RoboDK station: Conveyor_Station.rdk

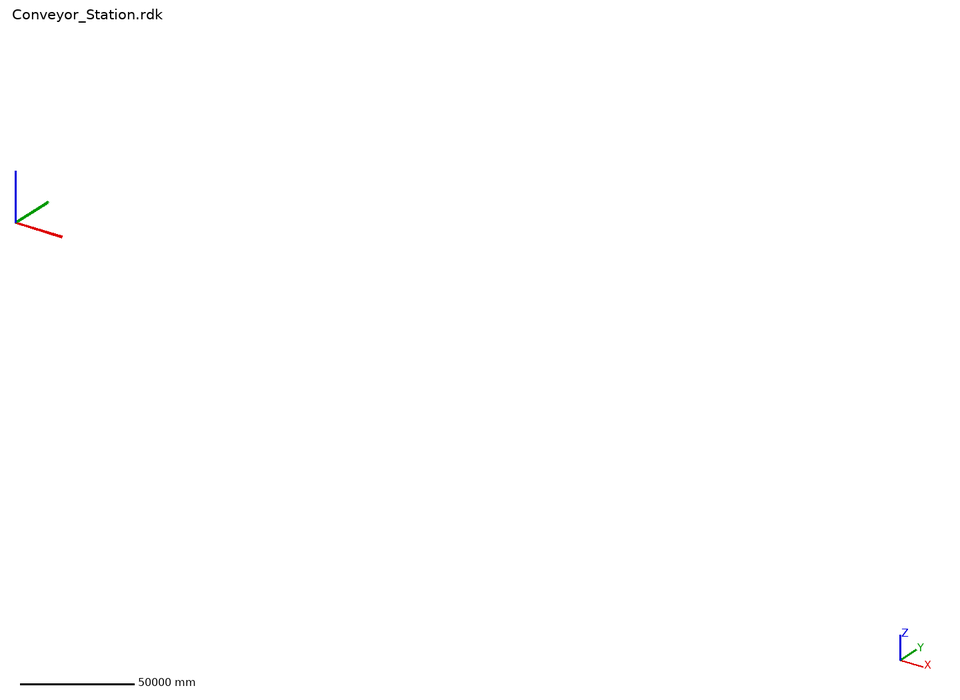
[picture v0: the station drawn from its stored meshes, robots at their saved joint values, targets as dots, program paths as lines]
Station Conveyor_Station (saved by RoboDK 6.0.1). Poses are relative to the parent item; angles as X-Y-Z fixed-axis rotations.
  - frame Conveyor Belt Wide (2m) Base at (0, 0, 0) mm
    - robot Conveyor Belt Wide (2m): 1 axes
        modified DH rows (alpha deg, a mm, theta deg, d mm): 0, 0, 0, 0 linear
        base shift (0, 0, 0) mm, rotated rx 0 ry 90 rz 0 deg
        joint limits [-900000] to [900000]; home [0]; saved at [-400005]
      - frame Conveyor Frame at (0, 0, 0) mm
        - object Box at (896234, 103.35, 13.17) mm, rotated rx -0.5 ry 0.31 rz 13.64 deg, size 10 x 20 x 5 mm, geometry from box.sld
        - object Box at (895766, 103.35, 13.17) mm, rotated rx -0.51 ry 0.3 rz 12.18 deg, size 10 x 20 x 5 mm, geometry from box.sld
        - object Box at (895300, 103.35, 13.17) mm, rotated rx -0.59 ry -0.09 rz -27.08 deg, size 10 x 20 x 5 mm, geometry from box.sld
        - object Box at (894830, 103.35, 13.17) mm, rotated rx -0.59 ry 0.03 rz -14.87 deg, size 10 x 20 x 5 mm, geometry from box.sld
        - object Box at (894363, 103.35, 13.17) mm, rotated rx -0.59 ry 0.08 rz -10.87 deg, size 10 x 20 x 5 mm, geometry from box.sld
        - object Box at (893893, 103.35, 13.17) mm, rotated rx -0.54 ry -0.25 rz -42.71 deg, size 10 x 20 x 5 mm, geometry from box.sld
        - object Box at (893423, 103.35, 13.17) mm, rotated rx -0.58 ry -0.12 rz -29.69 deg, size 10 x 20 x 5 mm, geometry from box.sld
        - object Box at (892951, 103.35, 13.17) mm, rotated rx -0.54 ry -0.25 rz -42.74 deg, size 10 x 20 x 5 mm, geometry from box.sld
        - object Box at (892481, 103.35, 13.17) mm, rotated rx -0.56 ry -0.19 rz -36.39 deg, size 10 x 20 x 5 mm, geometry from box.sld
        - object Box at (892010, 103.35, 13.17) mm, rotated rx -0.38 ry 0.45 rz 31.55 deg, size 10 x 20 x 5 mm, geometry from box.sld
        - object Box at (891537, 103.35, 13.17) mm, rotated rx -0.58 ry -0.14 rz -31.84 deg, size 10 x 20 x 5 mm, geometry from box.sld
        - object Box at (891061, 103.35, 13.17) mm, rotated rx -0.45 ry 0.39 rz 23.02 deg, size 10 x 20 x 5 mm, geometry from box.sld
        - object Box at (889213, 103.35, 13.17) mm, rotated rx -0.58 ry 0.14 rz -4.6 deg, size 10 x 20 x 5 mm, geometry from box.sld
        - object Box at (887815, 103.35, 13.17) mm, rotated rx -0.5 ry 0.33 rz 15.16 deg, size 10 x 20 x 5 mm, geometry from box.sld
        - object Box at (884546, 103.35, 13.17) mm, rotated rx -0.51 ry 0.31 rz 13.23 deg, size 10 x 20 x 5 mm, geometry from box.sld
        - object Box at (884069, 103.35, 13.17) mm, rotated rx -0.53 ry -0.27 rz -44.95 deg, size 10 x 20 x 5 mm, geometry from box.sld
        - object Box at (883940, 103.35, 13.17) mm, rotated rx -0.42 ry 0.42 rz 26.41 deg, size 10 x 20 x 5 mm, geometry from box.sld
        - object Box at (883628, 103.35, 13.17) mm, rotated rx -0.43 ry 0.41 rz 25.46 deg, size 10 x 20 x 5 mm, geometry from box.sld
        - object Box at (881822, 103.35, 13.17) mm, rotated rx -0.29 ry 0.52 rz 42.29 deg, size 10 x 20 x 5 mm, geometry from box.sld
        - object Box at (881392, 103.35, 13.17) mm, rotated rx -0.58 ry 0.12 rz -6.43 deg, size 10 x 20 x 5 mm, geometry from box.sld
        - object Box at (880938, 103.35, 13.17) mm, rotated rx -0.33 ry 0.5 rz 38.54 deg, size 10 x 20 x 5 mm, geometry from box.sld
        - object Box at (880498, 103.35, 13.17) mm, rotated rx -0.44 ry 0.4 rz 23.86 deg, size 10 x 20 x 5 mm, geometry from box.sld
        - object Box at (880042, 103.35, 13.17) mm, rotated rx -0.58 ry 0.13 rz -5.68 deg, size 10 x 20 x 5 mm, geometry from box.sld
        - object Box at (879599, 103.35, 13.17) mm, rotated rx -0.55 ry 0.22 rz 3.99 deg, size 10 x 20 x 5 mm, geometry from box.sld
        - object Box at (879164, 103.35, 13.17) mm, rotated rx -0.59 ry -0.01 rz -18.88 deg, size 10 x 20 x 5 mm, geometry from box.sld
        - object Box at (878722, 103.35, 13.17) mm, rotated rx -0.54 ry -0.24 rz -41.68 deg, size 10 x 20 x 5 mm, geometry from box.sld
        - object Box at (878276, 103.35, 13.17) mm, rotated rx -0.43 ry 0.41 rz 25.6 deg, size 10 x 20 x 5 mm, geometry from box.sld
        - object Box at (877829, 103.35, 13.17) mm, rotated rx -0.55 ry 0.23 rz 4.27 deg, size 10 x 20 x 5 mm, geometry from box.sld
        - object Box at (877389, 103.35, 13.17) mm, rotated rx -0.49 ry 0.33 rz 16.13 deg, size 10 x 20 x 5 mm, geometry from box.sld
        - object Box at (876944, 103.35, 13.17) mm, rotated rx -0.5 ry 0.33 rz 15.3 deg, size 10 x 20 x 5 mm, geometry from box.sld
        - object Box at (876499, 103.35, 13.17) mm, rotated rx -0.33 ry 0.5 rz 38.6 deg, size 10 x 20 x 5 mm, geometry from box.sld
        - object Box at (876043, 103.35, 13.17) mm, rotated rx -0.41 ry 0.43 rz 28.42 deg, size 10 x 20 x 5 mm, geometry from box.sld
        - object Box at (875592, 103.35, 13.17) mm, rotated rx -0.59 ry 0.03 rz -15.71 deg, size 10 x 20 x 5 mm, geometry from box.sld
        - object Box at (867999, 103.35, 13.17) mm, rotated rx -0.55 ry -0.22 rz -39.96 deg, size 10 x 20 x 5 mm, geometry from box.sld
        - object Box at (867540, 103.35, 13.17) mm, rotated rx -0.43 ry 0.41 rz 25.54 deg, size 10 x 20 x 5 mm, geometry from box.sld
        - object Box at (867083, 103.35, 13.17) mm, rotated rx -0.55 ry 0.23 rz 5.04 deg, size 10 x 20 x 5 mm, geometry from box.sld
        - object Box at (866626, 103.35, 13.17) mm, rotated rx -0.53 ry 0.26 rz 7.77 deg, size 10 x 20 x 5 mm, geometry from box.sld
        - object Box at (866172, 103.35, 13.17) mm, rotated rx -0.59 ry 0.09 rz -9.75 deg, size 10 x 20 x 5 mm, geometry from box.sld
        - object Box at (865727, 103.35, 13.17) mm, rotated rx -0.51 ry 0.31 rz 13.25 deg, size 10 x 20 x 5 mm, geometry from box.sld
        - object Box at (865279, 103.35, 13.17) mm, rotated rx -0.54 ry 0.24 rz 5.36 deg, size 10 x 20 x 5 mm, geometry from box.sld
        - object Box at (864826, 103.35, 13.17) mm, rotated rx -0.55 ry 0.23 rz 4.39 deg, size 10 x 20 x 5 mm, geometry from box.sld
        - object Box at (864371, 103.35, 13.17) mm, rotated rx -0.4 ry 0.44 rz 29 deg, size 10 x 20 x 5 mm, geometry from box.sld
        - object Box at (863914, 103.35, 13.17) mm, rotated rx -0.59 ry 0.09 rz -9.63 deg, size 10 x 20 x 5 mm, geometry from box.sld
        - object Box at (863455, 103.35, 13.17) mm, rotated rx -0.55 ry -0.22 rz -39.93 deg, size 10 x 20 x 5 mm, geometry from box.sld
        - object Box at (862988, 103.35, 13.17) mm, rotated rx -0.37 ry 0.46 rz 33.18 deg, size 10 x 20 x 5 mm, geometry from box.sld
        - object Box at (862512, 103.35, 13.17) mm, rotated rx -0.42 ry 0.42 rz 26.7 deg, size 10 x 20 x 5 mm, geometry from box.sld
        - object Box at (862049, 103.35, 13.17) mm, rotated rx -0.59 ry -0.07 rz -25.35 deg, size 10 x 20 x 5 mm, geometry from box.sld
        - object Box at (861585, 103.35, 13.17) mm, rotated rx -0.58 ry -0.13 rz -30.37 deg, size 10 x 20 x 5 mm, geometry from box.sld
        - object Box at (861121, 103.35, 13.17) mm, rotated rx -0.48 ry 0.35 rz 17.4 deg, size 10 x 20 x 5 mm, geometry from box.sld
        - object Box at (860654, 103.35, 13.17) mm, rotated rx -0.3 ry 0.51 rz 41.14 deg, size 10 x 20 x 5 mm, geometry from box.sld
        - object Box at (860190, 103.35, 13.17) mm, rotated rx -0.56 ry 0.2 rz 1.9 deg, size 10 x 20 x 5 mm, geometry from box.sld
        - object Box at (859725, 103.35, 13.17) mm, rotated rx -0.56 ry -0.21 rz -38.78 deg, size 10 x 20 x 5 mm, geometry from box.sld
        - object Box at (859255, 103.35, 13.17) mm, rotated rx -0.54 ry -0.25 rz -42.79 deg, size 10 x 20 x 5 mm, geometry from box.sld
        - object Box at (858791, 103.35, 13.17) mm, rotated rx -0.45 ry 0.38 rz 21.87 deg, size 10 x 20 x 5 mm, geometry from box.sld
        - object Box at (858319, 103.35, 13.17) mm, rotated rx -0.56 ry -0.21 rz -38.56 deg, size 10 x 20 x 5 mm, geometry from box.sld
        - object Box at (857850, 103.35, 13.17) mm, rotated rx -0.59 ry 0.09 rz -9.73 deg, size 10 x 20 x 5 mm, geometry from box.sld
        - object Box at (857380, 103.35, 13.17) mm, rotated rx -0.51 ry 0.31 rz 13.08 deg, size 10 x 20 x 5 mm, geometry from box.sld
        - object Box at (856914, 103.35, 13.17) mm, rotated rx -0.57 ry 0.16 rz -2.36 deg, size 10 x 20 x 5 mm, geometry from box.sld
        - object Box at (856441, 103.35, 13.17) mm, rotated rx -0.55 ry 0.23 rz 4.5 deg, size 10 x 20 x 5 mm, geometry from box.sld
        - object Box at (855972, 103.35, 13.17) mm, rotated rx -0.58 ry 0.13 rz -5.45 deg, size 10 x 20 x 5 mm, geometry from box.sld
        - object Box at (855499, 103.35, 13.17) mm, rotated rx -0.28 ry 0.52 rz 43.43 deg, size 10 x 20 x 5 mm, geometry from box.sld
        - object Box at (855027, 103.35, 13.17) mm, rotated rx -0.54 ry -0.24 rz -42.08 deg, size 10 x 20 x 5 mm, geometry from box.sld
        - object Box at (854558, 103.35, 13.17) mm, rotated rx -0.58 ry -0.12 rz -30.27 deg, size 10 x 20 x 5 mm, geometry from box.sld
        - object Box at (854093, 103.35, 13.17) mm, rotated rx -0.46 ry 0.37 rz 20.93 deg, size 10 x 20 x 5 mm, geometry from box.sld
        - object Box at (853622, 103.35, 13.17) mm, rotated rx -0.55 ry 0.23 rz 4.81 deg, size 10 x 20 x 5 mm, geometry from box.sld
        - object Box at (853148, 103.35, 13.17) mm, rotated rx -0.4 ry 0.44 rz 29.12 deg, size 10 x 20 x 5 mm, geometry from box.sld
        - object Box at (852676, 103.35, 13.17) mm, rotated rx -0.58 ry 0.14 rz -4.4 deg, size 10 x 20 x 5 mm, geometry from box.sld
        - object Box at (852209, 103.35, 13.17) mm, rotated rx -0.55 ry -0.22 rz -39.44 deg, size 10 x 20 x 5 mm, geometry from box.sld
        - object Box at (851737, 103.35, 13.17) mm, rotated rx -0.48 ry 0.35 rz 18.04 deg, size 10 x 20 x 5 mm, geometry from box.sld
        - object Box at (851258, 103.35, 13.17) mm, rotated rx -0.56 ry 0.2 rz 1.49 deg, size 10 x 20 x 5 mm, geometry from box.sld
        - object Box at (850779, 103.35, 13.17) mm, rotated rx -0.59 ry -0.05 rz -22.99 deg, size 10 x 20 x 5 mm, geometry from box.sld
        - object Box at (850302, 103.35, 13.17) mm, rotated rx -0.58 ry -0.14 rz -32.02 deg, size 10 x 20 x 5 mm, geometry from box.sld
        - object Box at (849825, 103.35, 13.17) mm, rotated rx -0.53 ry 0.27 rz 9.09 deg, size 10 x 20 x 5 mm, geometry from box.sld
        - object Box at (849347, 103.35, 13.17) mm, rotated rx -0.58 ry 0.1 rz -8 deg, size 10 x 20 x 5 mm, geometry from box.sld
        - object Box at (848871, 103.35, 13.17) mm, rotated rx -0.29 ry 0.52 rz 42.76 deg, size 10 x 20 x 5 mm, geometry from box.sld
        - object Box at (848385, 103.35, 13.17) mm, rotated rx -0.32 ry 0.5 rz 39.44 deg, size 10 x 20 x 5 mm, geometry from box.sld
        - object Box at (847911, 103.35, 13.17) mm, rotated rx -0.54 ry 0.24 rz 6.18 deg, size 10 x 20 x 5 mm, geometry from box.sld
        - object Box at (847434, 103.35, 13.17) mm, rotated rx -0.53 ry 0.27 rz 8.37 deg, size 10 x 20 x 5 mm, geometry from box.sld
        - object Box at (846952, 103.35, 13.17) mm, rotated rx -0.55 ry 0.21 rz 2.67 deg, size 10 x 20 x 5 mm, geometry from box.sld
        - object Box at (846476, 103.35, 13.17) mm, rotated rx -0.47 ry 0.36 rz 19.66 deg, size 10 x 20 x 5 mm, geometry from box.sld
        - object Box at (845998, 103.35, 13.17) mm, rotated rx -0.32 ry 0.5 rz 39.15 deg, size 10 x 20 x 5 mm, geometry from box.sld
        - object Box at (845516, 103.35, 13.17) mm, rotated rx -0.57 ry 0.18 rz -0.46 deg, size 10 x 20 x 5 mm, geometry from box.sld
        - object Box at (845034, 103.35, 13.17) mm, rotated rx -0.59 ry -0.04 rz -21.91 deg, size 10 x 20 x 5 mm, geometry from box.sld
        - object Box at (844553, 103.35, 13.17) mm, rotated rx -0.59 ry -0.09 rz -26.83 deg, size 10 x 20 x 5 mm, geometry from box.sld
        - object Box at (844070, 103.35, 13.17) mm, rotated rx -0.59 ry -0.01 rz -19.02 deg, size 10 x 20 x 5 mm, geometry from box.sld
        - object Box at (843586, 103.35, 13.17) mm, rotated rx -0.59 ry -0.08 rz -25.81 deg, size 10 x 20 x 5 mm, geometry from box.sld
        - object Box at (843104, 103.35, 13.17) mm, rotated rx -0.59 ry -0.01 rz -19.6 deg, size 10 x 20 x 5 mm, geometry from box.sld
        - object Box at (842621, 103.35, 13.17) mm, rotated rx -0.38 ry 0.45 rz 31.78 deg, size 10 x 20 x 5 mm, geometry from box.sld
        - object Box at (842135, 103.35, 13.17) mm, rotated rx -0.55 ry -0.23 rz -40.91 deg, size 10 x 20 x 5 mm, geometry from box.sld
        - object Box at (841652, 103.35, 13.17) mm, rotated rx -0.59 ry -0.05 rz -22.69 deg, size 10 x 20 x 5 mm, geometry from box.sld
        - object Box at (841168, 103.35, 13.17) mm, rotated rx -0.54 ry -0.26 rz -43.77 deg, size 10 x 20 x 5 mm, geometry from box.sld
        - object Box at (840683, 103.35, 13.17) mm, rotated rx -0.39 ry 0.45 rz 30.57 deg, size 10 x 20 x 5 mm, geometry from box.sld
        - object Box at (840198, 103.35, 13.17) mm, rotated rx -0.57 ry -0.16 rz -33.5 deg, size 10 x 20 x 5 mm, geometry from box.sld
        - object Box at (839715, 103.35, 13.17) mm, rotated rx -0.58 ry -0.12 rz -30.28 deg, size 10 x 20 x 5 mm, geometry from box.sld
        - object Box at (839227, 103.35, 13.17) mm, rotated rx -0.35 ry 0.48 rz 35.52 deg, size 10 x 20 x 5 mm, geometry from box.sld
        - object Box at (838741, 103.35, 13.17) mm, rotated rx -0.58 ry 0.1 rz -8.02 deg, size 10 x 20 x 5 mm, geometry from box.sld
        - object Box at (838251, 103.35, 13.17) mm, rotated rx -0.57 ry -0.15 rz -33.01 deg, size 10 x 20 x 5 mm, geometry from box.sld
        - object Box at (837766, 103.35, 13.17) mm, rotated rx -0.47 ry 0.36 rz 19.31 deg, size 10 x 20 x 5 mm, geometry from box.sld
        - object Box at (837279, 103.35, 13.17) mm, rotated rx -0.57 ry 0.15 rz -3.62 deg, size 10 x 20 x 5 mm, geometry from box.sld
        - object Box at (836786, 103.35, 13.17) mm, rotated rx -0.3 ry 0.51 rz 41.2 deg, size 10 x 20 x 5 mm, geometry from box.sld
        - object Box at (836295, 103.35, 13.17) mm, rotated rx -0.35 ry 0.48 rz 35.79 deg, size 10 x 20 x 5 mm, geometry from box.sld
        - object Box at (835805, 103.35, 13.17) mm, rotated rx -0.58 ry 0.11 rz -7.26 deg, size 10 x 20 x 5 mm, geometry from box.sld
        - object Box at (835317, 103.35, 13.17) mm, rotated rx -0.58 ry 0.14 rz -4.75 deg, size 10 x 20 x 5 mm, geometry from box.sld
        - object Box at (834829, 103.35, 13.17) mm, rotated rx -0.48 ry 0.35 rz 18.31 deg, size 10 x 20 x 5 mm, geometry from box.sld
        - object Box at (834338, 103.35, 13.17) mm, rotated rx -0.44 ry 0.4 rz 24.11 deg, size 10 x 20 x 5 mm, geometry from box.sld
        - object Box at (833842, 103.35, 13.17) mm, rotated rx -0.55 ry -0.22 rz -39.64 deg, size 10 x 20 x 5 mm, geometry from box.sld
        - object Box at (833349, 103.35, 13.17) mm, rotated rx -0.46 ry 0.37 rz 20.57 deg, size 10 x 20 x 5 mm, geometry from box.sld
        - object Box at (832860, 103.35, 13.17) mm, rotated rx -0.55 ry -0.23 rz -40.82 deg, size 10 x 20 x 5 mm, geometry from box.sld
        - object Box at (832363, 103.35, 13.17) mm, rotated rx -0.58 ry 0.1 rz -8.13 deg, size 10 x 20 x 5 mm, geometry from box.sld
        - object Box at (831873, 103.35, 13.17) mm, rotated rx -0.59 ry -0.08 rz -26.3 deg, size 10 x 20 x 5 mm, geometry from box.sld
        - object Box at (831377, 103.35, 13.17) mm, rotated rx -0.52 ry 0.28 rz 10.12 deg, size 10 x 20 x 5 mm, geometry from box.sld
        - object Box at (830887, 103.35, 13.17) mm, rotated rx -0.59 ry 0.02 rz -16.15 deg, size 10 x 20 x 5 mm, geometry from box.sld
        - object Box at (830394, 103.35, 13.17) mm, rotated rx -0.59 ry -0.03 rz -21.06 deg, size 10 x 20 x 5 mm, geometry from box.sld
        - object Box at (829901, 103.35, 13.17) mm, rotated rx -0.59 ry -0.02 rz -20.25 deg, size 10 x 20 x 5 mm, geometry from box.sld
        - object Box at (829404, 103.35, 13.17) mm, rotated rx -0.49 ry 0.34 rz 17.03 deg, size 10 x 20 x 5 mm, geometry from box.sld
        - object Box at (828911, 103.35, 13.17) mm, rotated rx -0.56 ry 0.19 rz 0.53 deg, size 10 x 20 x 5 mm, geometry from box.sld
        - object Box at (828417, 103.35, 13.17) mm, rotated rx -0.32 ry 0.5 rz 38.99 deg, size 10 x 20 x 5 mm, geometry from box.sld
        - object Box at (827919, 103.35, 13.17) mm, rotated rx -0.58 ry -0.14 rz -31.79 deg, size 10 x 20 x 5 mm, geometry from box.sld
        - object Box at (827419, 103.35, 13.17) mm, rotated rx -0.47 ry 0.36 rz 19.71 deg, size 10 x 20 x 5 mm, geometry from box.sld
        - object Box at (826919, 103.35, 13.17) mm, rotated rx -0.28 ry 0.52 rz 43.35 deg, size 10 x 20 x 5 mm, geometry from box.sld
        - object Box at (826422, 103.35, 13.17) mm, rotated rx -0.47 ry 0.37 rz 20.05 deg, size 10 x 20 x 5 mm, geometry from box.sld
        - object Box at (825923, 103.35, 13.17) mm, rotated rx -0.59 ry -0.09 rz -27.23 deg, size 10 x 20 x 5 mm, geometry from box.sld
        - object Box at (825422, 103.35, 13.17) mm, rotated rx -0.59 ry -0.02 rz -20.55 deg, size 10 x 20 x 5 mm, geometry from box.sld
        - object Box at (824929, 103.35, 13.17) mm, rotated rx -0.54 ry 0.25 rz 6.23 deg, size 10 x 20 x 5 mm, geometry from box.sld
        - object Box at (824425, 103.35, 13.17) mm, rotated rx -0.59 ry 0 rz -17.98 deg, size 10 x 20 x 5 mm, geometry from box.sld
        - object Box at (823928, 103.35, 13.17) mm, rotated rx -0.31 ry 0.5 rz 39.89 deg, size 10 x 20 x 5 mm, geometry from box.sld
        - object Box at (823424, 103.35, 13.17) mm, rotated rx -0.55 ry 0.23 rz 4.6 deg, size 10 x 20 x 5 mm, geometry from box.sld
        - object Box at (822920, 103.35, 13.17) mm, rotated rx -0.4 ry 0.44 rz 29.82 deg, size 10 x 20 x 5 mm, geometry from box.sld
        - object Box at (822418, 103.35, 13.17) mm, rotated rx -0.34 ry 0.49 rz 36.72 deg, size 10 x 20 x 5 mm, geometry from box.sld
        - object Box at (821917, 103.35, 13.17) mm, rotated rx -0.58 ry -0.12 rz -30.21 deg, size 10 x 20 x 5 mm, geometry from box.sld
        - object Box at (821420, 103.35, 13.17) mm, rotated rx -0.59 ry 0.04 rz -14.15 deg, size 10 x 20 x 5 mm, geometry from box.sld
        - object Box at (820919, 103.35, 13.17) mm, rotated rx -0.59 ry -0.08 rz -25.75 deg, size 10 x 20 x 5 mm, geometry from box.sld
        - object Box at (820410, 103.35, 13.17) mm, rotated rx -0.5 ry 0.33 rz 15.32 deg, size 10 x 20 x 5 mm, geometry from box.sld
        - object Box at (819909, 103.35, 13.17) mm, rotated rx -0.53 ry 0.26 rz 7.55 deg, size 10 x 20 x 5 mm, geometry from box.sld
        - object Box at (819403, 103.35, 13.17) mm, rotated rx -0.28 ry 0.52 rz 43.76 deg, size 10 x 20 x 5 mm, geometry from box.sld
        - object Box at (818898, 103.35, 13.17) mm, rotated rx -0.55 ry 0.21 rz 2.65 deg, size 10 x 20 x 5 mm, geometry from box.sld
        - object Box at (818392, 103.35, 13.17) mm, rotated rx -0.32 ry 0.5 rz 39.41 deg, size 10 x 20 x 5 mm, geometry from box.sld
        - object Box at (817887, 103.35, 13.17) mm, rotated rx -0.33 ry 0.49 rz 38.25 deg, size 10 x 20 x 5 mm, geometry from box.sld
        - object Box at (817383, 103.35, 13.17) mm, rotated rx -0.58 ry -0.11 rz -28.6 deg, size 10 x 20 x 5 mm, geometry from box.sld
        - object Box at (816879, 103.35, 13.17) mm, rotated rx -0.38 ry 0.46 rz 31.95 deg, size 10 x 20 x 5 mm, geometry from box.sld
        - object Box at (816374, 103.35, 13.17) mm, rotated rx -0.3 ry 0.51 rz 41.87 deg, size 10 x 20 x 5 mm, geometry from box.sld
        - object Box at (815868, 103.35, 13.17) mm, rotated rx -0.28 ry 0.52 rz 44.01 deg, size 10 x 20 x 5 mm, geometry from box.sld
        - object Box at (815360, 103.35, 13.17) mm, rotated rx -0.37 ry 0.46 rz 32.8 deg, size 10 x 20 x 5 mm, geometry from box.sld
        - object Box at (814853, 103.35, 13.17) mm, rotated rx -0.59 ry 0.07 rz -11.65 deg, size 10 x 20 x 5 mm, geometry from box.sld
        - object Box at (814348, 103.35, 13.17) mm, rotated rx -0.59 ry 0 rz -18.55 deg, size 10 x 20 x 5 mm, geometry from box.sld
        - object Box at (813832, 103.35, 13.17) mm, rotated rx -0.44 ry 0.4 rz 24.43 deg, size 10 x 20 x 5 mm, geometry from box.sld
        - object Box at (813321, 103.35, 13.17) mm, rotated rx -0.51 ry 0.31 rz 13.24 deg, size 10 x 20 x 5 mm, geometry from box.sld
        - object Box at (812812, 103.35, 13.17) mm, rotated rx -0.41 ry 0.43 rz 28.3 deg, size 10 x 20 x 5 mm, geometry from box.sld
        - object Box at (812298, 103.35, 13.17) mm, rotated rx -0.27 ry 0.53 rz 44.37 deg, size 10 x 20 x 5 mm, geometry from box.sld
        - object Box at (811784, 103.35, 13.17) mm, rotated rx -0.5 ry 0.32 rz 13.91 deg, size 10 x 20 x 5 mm, geometry from box.sld
        - object Box at (811274, 103.35, 13.17) mm, rotated rx -0.59 ry -0.02 rz -20.03 deg, size 10 x 20 x 5 mm, geometry from box.sld
        - object Box at (810763, 103.35, 13.17) mm, rotated rx -0.59 ry -0.02 rz -19.79 deg, size 10 x 20 x 5 mm, geometry from box.sld
        - object Box at (810254, 103.35, 13.17) mm, rotated rx -0.35 ry 0.48 rz 35.74 deg, size 10 x 20 x 5 mm, geometry from box.sld
        - object Box at (809736, 103.35, 13.17) mm, rotated rx -0.59 ry 0.09 rz -9.12 deg, size 10 x 20 x 5 mm, geometry from box.sld
        - object Box at (809227, 103.35, 13.17) mm, rotated rx -0.56 ry 0.19 rz 0.29 deg, size 10 x 20 x 5 mm, geometry from box.sld
        - object Box at (808709, 103.35, 13.17) mm, rotated rx -0.38 ry 0.45 rz 31.82 deg, size 10 x 20 x 5 mm, geometry from box.sld
        - object Box at (808195, 103.35, 13.17) mm, rotated rx -0.4 ry 0.44 rz 29.46 deg, size 10 x 20 x 5 mm, geometry from box.sld
        - object Box at (807680, 103.35, 13.17) mm, rotated rx -0.53 ry 0.26 rz 7.88 deg, size 10 x 20 x 5 mm, geometry from box.sld
        - object Box at (807162, 103.35, 13.17) mm, rotated rx -0.51 ry 0.3 rz 12.3 deg, size 10 x 20 x 5 mm, geometry from box.sld
        - object Box at (806641, 103.35, 13.17) mm, rotated rx -0.3 ry 0.51 rz 41.63 deg, size 10 x 20 x 5 mm, geometry from box.sld
        - object Box at (806130, 103.35, 13.17) mm, rotated rx -0.56 ry 0.19 rz 0.61 deg, size 10 x 20 x 5 mm, geometry from box.sld
        - object Box at (805613, 103.35, 13.17) mm, rotated rx -0.45 ry 0.39 rz 22.73 deg, size 10 x 20 x 5 mm, geometry from box.sld
        - object Box at (805094, 103.35, 13.17) mm, rotated rx -0.59 ry -0.03 rz -20.82 deg, size 10 x 20 x 5 mm, geometry from box.sld
        - object Box at (804579, 103.35, 13.17) mm, rotated rx -0.55 ry -0.22 rz -40.13 deg, size 10 x 20 x 5 mm, geometry from box.sld
        - object Box at (804064, 103.35, 13.17) mm, rotated rx -0.58 ry 0.13 rz -5.18 deg, size 10 x 20 x 5 mm, geometry from box.sld
        - object Box at (803548, 103.35, 13.17) mm, rotated rx -0.55 ry 0.21 rz 2.72 deg, size 10 x 20 x 5 mm, geometry from box.sld
        - object Box at (803030, 103.35, 13.17) mm, rotated rx -0.36 ry 0.47 rz 34.01 deg, size 10 x 20 x 5 mm, geometry from box.sld
        - object Box at (802512, 103.35, 13.17) mm, rotated rx -0.51 ry 0.3 rz 11.68 deg, size 10 x 20 x 5 mm, geometry from box.sld
        - object Box at (801994, 103.35, 13.17) mm, rotated rx -0.57 ry -0.17 rz -34.33 deg, size 10 x 20 x 5 mm, geometry from box.sld
        - object Box at (801472, 103.35, 13.17) mm, rotated rx -0.5 ry 0.32 rz 14.1 deg, size 10 x 20 x 5 mm, geometry from box.sld
        - object Box at (800951, 103.35, 13.17) mm, rotated rx -0.51 ry 0.31 rz 13.06 deg, size 10 x 20 x 5 mm, geometry from box.sld
        - object Box at (800432, 103.35, 13.17) mm, rotated rx -0.59 ry -0.02 rz -20.34 deg, size 10 x 20 x 5 mm, geometry from box.sld
        - object Box at (800001, 103.35, 13.17) mm, rotated rx -0.59 ry 0.03 rz -15.33 deg, size 10 x 20 x 5 mm, geometry from box.sld
        - object Box at (799501, 103.35, 13.17) mm, rotated rx -0.54 ry -0.25 rz -43.39 deg, size 10 x 20 x 5 mm, geometry from box.sld
        - object Box at (798979, 103.35, 13.17) mm, rotated rx -0.4 ry 0.44 rz 29.43 deg, size 10 x 20 x 5 mm, geometry from box.sld
        - object Box at (798451, 103.35, 13.17) mm, rotated rx -0.58 ry -0.13 rz -30.77 deg, size 10 x 20 x 5 mm, geometry from box.sld
        - object Box at (797933, 103.35, 13.17) mm, rotated rx -0.55 ry -0.21 rz -39.14 deg, size 10 x 20 x 5 mm, geometry from box.sld
        - object Box at (797410, 103.35, 13.17) mm, rotated rx -0.54 ry -0.24 rz -41.85 deg, size 10 x 20 x 5 mm, geometry from box.sld
        - object Box at (796890, 103.35, 13.17) mm, rotated rx -0.57 ry -0.17 rz -34.8 deg, size 10 x 20 x 5 mm, geometry from box.sld
        - object Box at (796360, 103.35, 13.17) mm, rotated rx -0.43 ry 0.41 rz 25.65 deg, size 10 x 20 x 5 mm, geometry from box.sld
        - object Box at (795838, 103.35, 13.17) mm, rotated rx -0.59 ry -0.09 rz -26.89 deg, size 10 x 20 x 5 mm, geometry from box.sld
        - object Box at (795317, 103.35, 13.17) mm, rotated rx -0.42 ry 0.42 rz 26.96 deg, size 10 x 20 x 5 mm, geometry from box.sld
        - object Box at (794795, 103.35, 13.17) mm, rotated rx -0.55 ry -0.22 rz -39.88 deg, size 10 x 20 x 5 mm, geometry from box.sld
        - object Box at (794268, 103.35, 13.17) mm, rotated rx -0.59 ry -0.01 rz -19.47 deg, size 10 x 20 x 5 mm, geometry from box.sld
        - object Box at (793735, 103.35, 13.17) mm, rotated rx -0.56 ry 0.2 rz 1.5 deg, size 10 x 20 x 5 mm, geometry from box.sld
        - object Box at (793205, 103.35, 13.17) mm, rotated rx -0.56 ry 0.19 rz 0.8 deg, size 10 x 20 x 5 mm, geometry from box.sld
        - object Box at (791620, 103.35, 13.17) mm, rotated rx -0.5 ry 0.32 rz 14.93 deg, size 10 x 20 x 5 mm, geometry from box.sld
        - object Box at (790003, 103.35, 13.17) mm, rotated rx -0.59 ry 0.01 rz -17.46 deg, size 10 x 20 x 5 mm, geometry from box.sld
        - object Box at (789472, 103.35, 13.17) mm, rotated rx -0.47 ry 0.37 rz 19.97 deg, size 10 x 20 x 5 mm, geometry from box.sld
        - object Box at (788941, 103.35, 13.17) mm, rotated rx -0.59 ry -0.02 rz -19.81 deg, size 10 x 20 x 5 mm, geometry from box.sld
        - object Box at (788418, 103.35, 13.17) mm, rotated rx -0.59 ry -0.02 rz -20.48 deg, size 10 x 20 x 5 mm, geometry from box.sld
        - object Box at (787893, 103.35, 13.17) mm, rotated rx -0.59 ry -0.08 rz -25.44 deg, size 10 x 20 x 5 mm, geometry from box.sld
        - object Box at (787376, 103.35, 13.17) mm, rotated rx -0.29 ry 0.52 rz 42.24 deg, size 10 x 20 x 5 mm, geometry from box.sld
        - object Box at (785262, 103.35, 13.17) mm, rotated rx -0.34 ry 0.48 rz 36.37 deg, size 10 x 20 x 5 mm, geometry from box.sld
        - object Box at (784703, 103.35, 13.17) mm, rotated rx -0.31 ry 0.51 rz 40.65 deg, size 10 x 20 x 5 mm, geometry from box.sld
        - object Box at (784140, 103.35, 13.17) mm, rotated rx -0.59 ry 0.02 rz -16.67 deg, size 10 x 20 x 5 mm, geometry from box.sld
        - object Box at (783610, 103.35, 13.17) mm, rotated rx -0.4 ry 0.44 rz 29.43 deg, size 10 x 20 x 5 mm, geometry from box.sld
        - object Box at (783080, 103.35, 13.17) mm, rotated rx -0.58 ry -0.14 rz -31.4 deg, size 10 x 20 x 5 mm, geometry from box.sld
        - object Box at (782548, 103.35, 13.17) mm, rotated rx -0.59 ry 0 rz -18.46 deg, size 10 x 20 x 5 mm, geometry from box.sld
        - object Box at (782009, 103.35, 13.17) mm, rotated rx -0.55 ry -0.22 rz -39.9 deg, size 10 x 20 x 5 mm, geometry from box.sld
        - object Box at (781485, 103.35, 13.17) mm, rotated rx -0.54 ry 0.24 rz 5.81 deg, size 10 x 20 x 5 mm, geometry from box.sld
        - object Box at (780962, 103.35, 13.17) mm, rotated rx -0.59 ry 0.06 rz -12.4 deg, size 10 x 20 x 5 mm, geometry from box.sld
        - object Box at (780427, 103.35, 13.17) mm, rotated rx -0.47 ry 0.37 rz 19.81 deg, size 10 x 20 x 5 mm, geometry from box.sld
        - object Box at (779895, 103.35, 13.17) mm, rotated rx -0.59 ry -0.07 rz -24.94 deg, size 10 x 20 x 5 mm, geometry from box.sld
        - object Box at (779360, 103.35, 13.17) mm, rotated rx -0.28 ry 0.52 rz 43.8 deg, size 10 x 20 x 5 mm, geometry from box.sld
        - object Box at (778825, 103.35, 13.17) mm, rotated rx -0.45 ry 0.39 rz 22.8 deg, size 10 x 20 x 5 mm, geometry from box.sld
        - object Box at (778291, 103.35, 13.17) mm, rotated rx -0.58 ry -0.14 rz -32.29 deg, size 10 x 20 x 5 mm, geometry from box.sld
        - object Box at (777770, 103.35, 13.17) mm, rotated rx -0.34 ry 0.49 rz 37.05 deg, size 10 x 20 x 5 mm, geometry from box.sld
        - object Box at (777234, 103.35, 13.17) mm, rotated rx -0.59 ry 0.08 rz -10.52 deg, size 10 x 20 x 5 mm, geometry from box.sld
        - object Box at (776677, 103.35, 13.17) mm, rotated rx -0.5 ry 0.32 rz 14.02 deg, size 10 x 20 x 5 mm, geometry from box.sld
        - object Box at (776136, 103.35, 13.17) mm, rotated rx -0.51 ry 0.31 rz 13.12 deg, size 10 x 20 x 5 mm, geometry from box.sld
        - object Box at (775600, 103.35, 13.17) mm, rotated rx -0.59 ry 0.1 rz -8.75 deg, size 10 x 20 x 5 mm, geometry from box.sld
        - object Box at (775057, 103.35, 13.17) mm, rotated rx -0.59 ry 0.07 rz -10.91 deg, size 10 x 20 x 5 mm, geometry from box.sld
        - object Box at (774530, 103.35, 13.17) mm, rotated rx -0.49 ry 0.34 rz 16.71 deg, size 10 x 20 x 5 mm, geometry from box.sld
        - object Box at (773989, 103.35, 13.17) mm, rotated rx -0.57 ry 0.15 rz -3.12 deg, size 10 x 20 x 5 mm, geometry from box.sld
        - object Box at (773453, 103.35, 13.17) mm, rotated rx -0.51 ry 0.31 rz 12.93 deg, size 10 x 20 x 5 mm, geometry from box.sld
        - object Box at (772909, 103.35, 13.17) mm, rotated rx -0.58 ry 0.12 rz -6.06 deg, size 10 x 20 x 5 mm, geometry from box.sld
        - object Box at (772376, 103.35, 13.17) mm, rotated rx -0.34 ry 0.49 rz 37.24 deg, size 10 x 20 x 5 mm, geometry from box.sld
        - object Box at (771828, 103.35, 13.17) mm, rotated rx -0.54 ry -0.25 rz -43.45 deg, size 10 x 20 x 5 mm, geometry from box.sld
        - object Box at (771292, 103.35, 13.17) mm, rotated rx -0.51 ry 0.31 rz 12.93 deg, size 10 x 20 x 5 mm, geometry from box.sld
        - object Box at (770765, 103.35, 13.17) mm, rotated rx -0.58 ry 0.12 rz -6.57 deg, size 10 x 20 x 5 mm, geometry from box.sld
        - object Box at (770213, 103.35, 13.17) mm, rotated rx -0.4 ry 0.44 rz 29.53 deg, size 10 x 20 x 5 mm, geometry from box.sld
        - object Box at (769672, 103.35, 13.17) mm, rotated rx -0.39 ry 0.45 rz 30.75 deg, size 10 x 20 x 5 mm, geometry from box.sld
        - object Box at (769131, 103.35, 13.17) mm, rotated rx -0.4 ry 0.44 rz 29.93 deg, size 10 x 20 x 5 mm, geometry from box.sld
        - object Box at (768601, 103.35, 13.17) mm, rotated rx -0.58 ry 0.1 rz -8.15 deg, size 10 x 20 x 5 mm, geometry from box.sld
        - object Box at (768056, 103.35, 13.17) mm, rotated rx -0.56 ry -0.19 rz -36.67 deg, size 10 x 20 x 5 mm, geometry from box.sld
        - object Box at (767497, 103.35, 13.17) mm, rotated rx -0.57 ry -0.16 rz -33.54 deg, size 10 x 20 x 5 mm, geometry from box.sld
        - object Box at (766950, 103.35, 13.17) mm, rotated rx -0.58 ry 0.14 rz -4.79 deg, size 10 x 20 x 5 mm, geometry from box.sld
        - object Box at (766411, 103.35, 13.17) mm, rotated rx -0.53 ry -0.26 rz -44.4 deg, size 10 x 20 x 5 mm, geometry from box.sld
        - object Box at (765869, 103.35, 13.17) mm, rotated rx -0.29 ry 0.52 rz 42.65 deg, size 10 x 20 x 5 mm, geometry from box.sld
        - object Box at (765328, 103.35, 13.17) mm, rotated rx -0.54 ry -0.24 rz -42.2 deg, size 10 x 20 x 5 mm, geometry from box.sld
        - object Box at (764778, 103.35, 13.17) mm, rotated rx -0.48 ry 0.35 rz 18.39 deg, size 10 x 20 x 5 mm, geometry from box.sld
        - object Box at (764237, 103.35, 13.17) mm, rotated rx -0.56 ry -0.2 rz -37.97 deg, size 10 x 20 x 5 mm, geometry from box.sld
        - object Box at (763694, 103.35, 13.17) mm, rotated rx -0.48 ry 0.35 rz 17.83 deg, size 10 x 20 x 5 mm, geometry from box.sld
        - object Box at (763136, 103.35, 13.17) mm, rotated rx -0.45 ry 0.39 rz 22.61 deg, size 10 x 20 x 5 mm, geometry from box.sld
        - object Box at (762576, 103.35, 13.17) mm, rotated rx -0.59 ry 0 rz -18.36 deg, size 10 x 20 x 5 mm, geometry from box.sld
        - object Box at (762042, 103.35, 13.17) mm, rotated rx -0.31 ry 0.51 rz 40.49 deg, size 10 x 20 x 5 mm, geometry from box.sld
        - object Box at (761489, 103.35, 13.17) mm, rotated rx -0.56 ry 0.2 rz 1.47 deg, size 10 x 20 x 5 mm, geometry from box.sld
        - object Box at (760946, 103.35, 13.17) mm, rotated rx -0.59 ry -0.09 rz -26.98 deg, size 10 x 20 x 5 mm, geometry from box.sld
        - object Box at (760411, 103.35, 13.17) mm, rotated rx -0.59 ry -0.06 rz -23.57 deg, size 10 x 20 x 5 mm, geometry from box.sld
        - object Box at (759851, 103.35, 13.17) mm, rotated rx -0.57 ry -0.17 rz -34.8 deg, size 10 x 20 x 5 mm, geometry from box.sld
        - object Box at (759238, 103.35, 13.17) mm, rotated rx -0.55 ry -0.23 rz -41.08 deg, size 10 x 20 x 5 mm, geometry from box.sld
        - object Box at (758681, 103.35, 13.17) mm, rotated rx -0.38 ry 0.46 rz 32.65 deg, size 10 x 20 x 5 mm, geometry from box.sld
        - object Box at (758134, 103.35, 13.17) mm, rotated rx -0.59 ry -0.03 rz -20.71 deg, size 10 x 20 x 5 mm, geometry from box.sld
        - object Box at (757567, 103.35, 13.17) mm, rotated rx -0.29 ry 0.52 rz 42.57 deg, size 10 x 20 x 5 mm, geometry from box.sld
        - object Box at (757016, 103.35, 13.17) mm, rotated rx -0.58 ry 0.11 rz -7.57 deg, size 10 x 20 x 5 mm, geometry from box.sld
        - object Box at (756466, 103.35, 13.17) mm, rotated rx -0.59 ry 0.03 rz -15.6 deg, size 10 x 20 x 5 mm, geometry from box.sld
        - object Box at (755922, 103.35, 13.17) mm, rotated rx -0.34 ry 0.48 rz 36.43 deg, size 10 x 20 x 5 mm, geometry from box.sld
        - object Box at (755365, 103.35, 13.17) mm, rotated rx -0.46 ry 0.37 rz 20.29 deg, size 10 x 20 x 5 mm, geometry from box.sld
        - object Box at (754794, 103.35, 13.17) mm, rotated rx -0.33 ry 0.49 rz 38.22 deg, size 10 x 20 x 5 mm, geometry from box.sld
        - object Box at (754238, 103.35, 13.17) mm, rotated rx -0.47 ry 0.36 rz 19.26 deg, size 10 x 20 x 5 mm, geometry from box.sld
        - object Box at (753693, 103.35, 13.17) mm, rotated rx -0.58 ry -0.12 rz -29.72 deg, size 10 x 20 x 5 mm, geometry from box.sld
        - object Box at (753143, 103.35, 13.17) mm, rotated rx -0.58 ry 0.15 rz -3.91 deg, size 10 x 20 x 5 mm, geometry from box.sld
        - object Box at (752591, 103.35, 13.17) mm, rotated rx -0.39 ry 0.45 rz 31.29 deg, size 10 x 20 x 5 mm, geometry from box.sld
        - object Box at (752035, 103.35, 13.17) mm, rotated rx -0.55 ry -0.22 rz -39.72 deg, size 10 x 20 x 5 mm, geometry from box.sld
        - object Box at (751485, 103.35, 13.17) mm, rotated rx -0.32 ry 0.5 rz 39.31 deg, size 10 x 20 x 5 mm, geometry from box.sld
        - object Box at (750924, 103.35, 13.17) mm, rotated rx -0.59 ry -0.03 rz -21.51 deg, size 10 x 20 x 5 mm, geometry from box.sld
        - object Box at (750360, 103.35, 13.17) mm, rotated rx -0.47 ry 0.36 rz 19.49 deg, size 10 x 20 x 5 mm, geometry from box.sld
        - object Box at (749800, 103.35, 13.17) mm, rotated rx -0.59 ry 0.08 rz -9.98 deg, size 10 x 20 x 5 mm, geometry from box.sld
        - object Box at (749232, 103.35, 13.17) mm, rotated rx -0.37 ry 0.46 rz 33.34 deg, size 10 x 20 x 5 mm, geometry from box.sld
        - object Box at (748682, 103.35, 13.17) mm, rotated rx -0.57 ry -0.15 rz -32.89 deg, size 10 x 20 x 5 mm, geometry from box.sld
        - object Box at (748124, 103.35, 13.17) mm, rotated rx -0.45 ry 0.39 rz 23.26 deg, size 10 x 20 x 5 mm, geometry from box.sld
        - object Box at (747566, 103.35, 13.17) mm, rotated rx -0.59 ry 0.1 rz -8.89 deg, size 10 x 20 x 5 mm, geometry from box.sld
        - object Box at (747036, 103.35, 13.17) mm, rotated rx -0.52 ry 0.3 rz 11.65 deg, size 10 x 20 x 5 mm, geometry from box.sld
        - object Box at (746459, 103.35, 13.17) mm, rotated rx -0.43 ry 0.41 rz 26.01 deg, size 10 x 20 x 5 mm, geometry from box.sld
        - object Box at (745902, 103.35, 13.17) mm, rotated rx -0.59 ry 0.03 rz -14.8 deg, size 10 x 20 x 5 mm, geometry from box.sld
        - object Box at (745342, 103.35, 13.17) mm, rotated rx -0.54 ry 0.25 rz 7 deg, size 10 x 20 x 5 mm, geometry from box.sld
        - object Box at (744781, 103.35, 13.17) mm, rotated rx -0.58 ry 0.11 rz -7.31 deg, size 10 x 20 x 5 mm, geometry from box.sld
        - object Box at (744212, 103.35, 13.17) mm, rotated rx -0.57 ry -0.16 rz -33.54 deg, size 10 x 20 x 5 mm, geometry from box.sld
        - object Box at (743652, 103.35, 13.17) mm, rotated rx -0.36 ry 0.47 rz 34.53 deg, size 10 x 20 x 5 mm, geometry from box.sld
        - object Box at (743080, 103.35, 13.17) mm, rotated rx -0.49 ry 0.34 rz 16.92 deg, size 10 x 20 x 5 mm, geometry from box.sld
        - object Box at (742503, 103.35, 13.17) mm, rotated rx -0.57 ry 0.16 rz -2.55 deg, size 10 x 20 x 5 mm, geometry from box.sld
        - object Box at (741946, 103.35, 13.17) mm, rotated rx -0.59 ry 0.08 rz -10 deg, size 10 x 20 x 5 mm, geometry from box.sld
        - object Box at (741382, 103.35, 13.17) mm, rotated rx -0.59 ry 0.06 rz -11.91 deg, size 10 x 20 x 5 mm, geometry from box.sld
        - object Box at (740819, 103.35, 13.17) mm, rotated rx -0.39 ry 0.45 rz 30.73 deg, size 10 x 20 x 5 mm, geometry from box.sld
        - object Box at (740247, 103.35, 13.17) mm, rotated rx -0.49 ry 0.34 rz 16.57 deg, size 10 x 20 x 5 mm, geometry from box.sld
        - object Box at (739684, 103.35, 13.17) mm, rotated rx -0.48 ry 0.35 rz 17.51 deg, size 10 x 20 x 5 mm, geometry from box.sld
        - object Box at (739114, 103.35, 13.17) mm, rotated rx -0.36 ry 0.47 rz 34.72 deg, size 10 x 20 x 5 mm, geometry from box.sld
        - object Box at (738552, 103.35, 13.17) mm, rotated rx -0.37 ry 0.47 rz 33.59 deg, size 10 x 20 x 5 mm, geometry from box.sld
        - object Box at (737996, 103.35, 13.17) mm, rotated rx -0.27 ry 0.53 rz 44.28 deg, size 10 x 20 x 5 mm, geometry from box.sld
        - object Box at (737399, 103.35, 13.17) mm, rotated rx -0.54 ry 0.25 rz 7.02 deg, size 10 x 20 x 5 mm, geometry from box.sld
        - object Box at (736827, 103.35, 13.17) mm, rotated rx -0.58 ry 0.12 rz -6.1 deg, size 10 x 20 x 5 mm, geometry from box.sld
        - object Box at (736253, 103.35, 13.17) mm, rotated rx -0.58 ry 0.14 rz -4.65 deg, size 10 x 20 x 5 mm, geometry from box.sld
        - object Box at (735678, 103.35, 13.17) mm, rotated rx -0.57 ry -0.17 rz -34.95 deg, size 10 x 20 x 5 mm, geometry from box.sld
        - object Box at (735106, 103.35, 13.17) mm, rotated rx -0.58 ry -0.1 rz -27.93 deg, size 10 x 20 x 5 mm, geometry from box.sld
        - object Box at (734539, 103.35, 13.17) mm, rotated rx -0.36 ry 0.47 rz 34.11 deg, size 10 x 20 x 5 mm, geometry from box.sld
        - object Box at (733962, 103.35, 13.17) mm, rotated rx -0.59 ry 0.09 rz -9.68 deg, size 10 x 20 x 5 mm, geometry from box.sld
        - object Box at (733396, 103.35, 13.17) mm, rotated rx -0.32 ry 0.5 rz 39.44 deg, size 10 x 20 x 5 mm, geometry from box.sld
        - object Box at (732826, 103.35, 13.17) mm, rotated rx -0.3 ry 0.51 rz 41.08 deg, size 10 x 20 x 5 mm, geometry from box.sld
        - object Box at (732252, 103.35, 13.17) mm, rotated rx -0.52 ry 0.29 rz 10.68 deg, size 10 x 20 x 5 mm, geometry from box.sld
        - object Box at (731692, 103.35, 13.17) mm, rotated rx -0.59 ry 0 rz -18.11 deg, size 10 x 20 x 5 mm, geometry from box.sld
        - object Box at (731106, 103.35, 13.17) mm, rotated rx -0.43 ry 0.41 rz 25.03 deg, size 10 x 20 x 5 mm, geometry from box.sld
        - object Box at (730548, 103.35, 13.17) mm, rotated rx -0.59 ry 0.06 rz -12.08 deg, size 10 x 20 x 5 mm, geometry from box.sld
        - object Box at (729974, 103.35, 13.17) mm, rotated rx -0.59 ry 0.04 rz -13.83 deg, size 10 x 20 x 5 mm, geometry from box.sld
        - object Box at (729390, 103.35, 13.17) mm, rotated rx -0.4 ry 0.44 rz 29.14 deg, size 10 x 20 x 5 mm, geometry from box.sld
        - object Box at (728813, 103.35, 13.17) mm, rotated rx -0.59 ry -0.02 rz -20.53 deg, size 10 x 20 x 5 mm, geometry from box.sld
        - object Box at (728245, 103.35, 13.17) mm, rotated rx -0.54 ry 0.25 rz 6.58 deg, size 10 x 20 x 5 mm, geometry from box.sld
        - object Box at (727671, 103.35, 13.17) mm, rotated rx -0.59 ry 0.07 rz -11.83 deg, size 10 x 20 x 5 mm, geometry from box.sld
        - object Box at (727097, 103.35, 13.17) mm, rotated rx -0.53 ry -0.26 rz -44.39 deg, size 10 x 20 x 5 mm, geometry from box.sld
        - object Box at (726521, 103.35, 13.17) mm, rotated rx -0.44 ry 0.4 rz 24.31 deg, size 10 x 20 x 5 mm, geometry from box.sld
        - object Box at (725947, 103.35, 13.17) mm, rotated rx -0.56 ry 0.19 rz 0.34 deg, size 10 x 20 x 5 mm, geometry from box.sld
        - object Box at (725372, 103.35, 13.17) mm, rotated rx -0.48 ry 0.35 rz 17.95 deg, size 10 x 20 x 5 mm, geometry from box.sld
        - object Box at (724774, 103.35, 13.17) mm, rotated rx -0.59 ry 0.09 rz -9.21 deg, size 10 x 20 x 5 mm, geometry from box.sld
        - object Box at (724199, 103.35, 13.17) mm, rotated rx -0.57 ry -0.16 rz -33.96 deg, size 10 x 20 x 5 mm, geometry from box.sld
        - object Box at (723621, 103.35, 13.17) mm, rotated rx -0.55 ry 0.24 rz 5.17 deg, size 10 x 20 x 5 mm, geometry from box.sld
        - object Box at (723049, 103.35, 13.17) mm, rotated rx -0.59 ry 0.01 rz -17.21 deg, size 10 x 20 x 5 mm, geometry from box.sld
        - object Box at (722458, 103.35, 13.17) mm, rotated rx -0.4 ry 0.44 rz 29.47 deg, size 10 x 20 x 5 mm, geometry from box.sld
        - object Box at (721880, 103.35, 13.17) mm, rotated rx -0.29 ry 0.52 rz 43.13 deg, size 10 x 20 x 5 mm, geometry from box.sld
        - object Box at (721284, 103.35, 13.17) mm, rotated rx -0.59 ry -0.01 rz -18.99 deg, size 10 x 20 x 5 mm, geometry from box.sld
        - object Box at (720699, 103.35, 13.17) mm, rotated rx -0.43 ry 0.41 rz 25.73 deg, size 10 x 20 x 5 mm, geometry from box.sld
        - object Box at (720121, 103.35, 13.17) mm, rotated rx -0.47 ry 0.36 rz 18.74 deg, size 10 x 20 x 5 mm, geometry from box.sld
        - object Box at (719536, 103.35, 13.17) mm, rotated rx -0.57 ry 0.17 rz -1.56 deg, size 10 x 20 x 5 mm, geometry from box.sld
        - object Box at (718948, 103.35, 13.17) mm, rotated rx -0.58 ry 0.12 rz -6.4 deg, size 10 x 20 x 5 mm, geometry from box.sld
        - object Box at (718360, 103.35, 13.17) mm, rotated rx -0.58 ry 0.13 rz -5.67 deg, size 10 x 20 x 5 mm, geometry from box.sld
        - object Box at (717766, 103.35, 13.17) mm, rotated rx -0.49 ry 0.33 rz 16.06 deg, size 10 x 20 x 5 mm, geometry from box.sld
        - object Box at (717166, 103.35, 13.17) mm, rotated rx -0.48 ry 0.35 rz 18.49 deg, size 10 x 20 x 5 mm, geometry from box.sld
        - object Box at (716596, 103.35, 13.17) mm, rotated rx -0.32 ry 0.5 rz 38.96 deg, size 10 x 20 x 5 mm, geometry from box.sld
        - object Box at (716011, 103.35, 13.17) mm, rotated rx -0.54 ry -0.24 rz -42.45 deg, size 10 x 20 x 5 mm, geometry from box.sld
        - object Box at (715428, 103.35, 13.17) mm, rotated rx -0.37 ry 0.47 rz 33.79 deg, size 10 x 20 x 5 mm, geometry from box.sld
        - object Box at (714834, 103.35, 13.17) mm, rotated rx -0.58 ry 0.14 rz -4.55 deg, size 10 x 20 x 5 mm, geometry from box.sld
        - object Box at (714234, 103.35, 13.17) mm, rotated rx -0.59 ry 0.06 rz -11.97 deg, size 10 x 20 x 5 mm, geometry from box.sld
        - object Box at (713642, 103.35, 13.17) mm, rotated rx -0.38 ry 0.45 rz 31.71 deg, size 10 x 20 x 5 mm, geometry from box.sld
        - object Box at (713043, 103.35, 13.17) mm, rotated rx -0.59 ry -0.07 rz -24.53 deg, size 10 x 20 x 5 mm, geometry from box.sld
        - object Box at (712454, 103.35, 13.17) mm, rotated rx -0.58 ry 0.11 rz -7.52 deg, size 10 x 20 x 5 mm, geometry from box.sld
        - object Box at (711876, 103.35, 13.17) mm, rotated rx -0.48 ry 0.35 rz 18.4 deg, size 10 x 20 x 5 mm, geometry from box.sld
        - object Box at (711289, 103.35, 13.17) mm, rotated rx -0.58 ry 0.13 rz -5.58 deg, size 10 x 20 x 5 mm, geometry from box.sld
        - object Box at (710705, 103.35, 13.17) mm, rotated rx -0.58 ry -0.12 rz -30.05 deg, size 10 x 20 x 5 mm, geometry from box.sld
        - object Box at (710097, 103.35, 13.17) mm, rotated rx -0.39 ry 0.44 rz 30.29 deg, size 10 x 20 x 5 mm, geometry from box.sld
        - object Box at (709492, 103.35, 13.17) mm, rotated rx -0.54 ry -0.25 rz -42.75 deg, size 10 x 20 x 5 mm, geometry from box.sld
        - object Box at (708907, 103.35, 13.17) mm, rotated rx -0.54 ry -0.24 rz -42.35 deg, size 10 x 20 x 5 mm, geometry from box.sld
        - object Box at (708314, 103.35, 13.17) mm, rotated rx -0.56 ry -0.19 rz -36.42 deg, size 10 x 20 x 5 mm, geometry from box.sld
        - object Box at (707715, 103.35, 13.17) mm, rotated rx -0.31 ry 0.51 rz 40.68 deg, size 10 x 20 x 5 mm, geometry from box.sld
        - object Box at (707117, 103.35, 13.17) mm, rotated rx -0.33 ry 0.49 rz 37.88 deg, size 10 x 20 x 5 mm, geometry from box.sld
        - object Box at (706518, 103.35, 13.17) mm, rotated rx -0.45 ry 0.39 rz 22.92 deg, size 10 x 20 x 5 mm, geometry from box.sld
        - object Box at (705907, 103.35, 13.17) mm, rotated rx -0.59 ry 0 rz -17.97 deg, size 10 x 20 x 5 mm, geometry from box.sld
        - object Box at (705314, 103.35, 13.17) mm, rotated rx -0.38 ry 0.46 rz 32.2 deg, size 10 x 20 x 5 mm, geometry from box.sld
        - object Box at (704729, 103.35, 13.17) mm, rotated rx -0.57 ry 0.16 rz -2.54 deg, size 10 x 20 x 5 mm, geometry from box.sld
        - object Box at (704146, 103.35, 13.17) mm, rotated rx -0.59 ry -0.09 rz -26.85 deg, size 10 x 20 x 5 mm, geometry from box.sld
        - object Box at (703551, 103.35, 13.17) mm, rotated rx -0.51 ry 0.3 rz 12.59 deg, size 10 x 20 x 5 mm, geometry from box.sld
        - object Box at (702970, 103.35, 13.17) mm, rotated rx -0.59 ry -0.03 rz -20.64 deg, size 10 x 20 x 5 mm, geometry from box.sld
        - object Box at (702349, 103.35, 13.17) mm, rotated rx -0.59 ry -0.03 rz -20.79 deg, size 10 x 20 x 5 mm, geometry from box.sld
        - object Box at (701739, 103.35, 13.17) mm, rotated rx -0.53 ry -0.26 rz -43.86 deg, size 10 x 20 x 5 mm, geometry from box.sld
        - object Box at (701147, 103.35, 13.17) mm, rotated rx -0.5 ry 0.31 rz 13.83 deg, size 10 x 20 x 5 mm, geometry from box.sld
        - object Box at (700540, 103.35, 13.17) mm, rotated rx -0.47 ry 0.36 rz 19.01 deg, size 10 x 20 x 5 mm, geometry from box.sld
        - object Box at (700002, 103.35, 13.17) mm, rotated rx -0.58 ry 0.12 rz -6.68 deg, size 10 x 20 x 5 mm, geometry from box.sld
        - object Box at (699789, 103.35, 13.17) mm, rotated rx -0.56 ry 0.19 rz 0.97 deg, size 10 x 20 x 5 mm, geometry from box.sld
        - object Box at (699197, 103.35, 13.17) mm, rotated rx -0.39 ry 0.44 rz 30.29 deg, size 10 x 20 x 5 mm, geometry from box.sld
        - object Box at (698577, 103.35, 13.17) mm, rotated rx -0.59 ry -0.06 rz -23.9 deg, size 10 x 20 x 5 mm, geometry from box.sld
        - object Box at (697976, 103.35, 13.17) mm, rotated rx -0.58 ry -0.11 rz -29.2 deg, size 10 x 20 x 5 mm, geometry from box.sld
        - object Box at (697374, 103.35, 13.17) mm, rotated rx -0.49 ry 0.33 rz 15.69 deg, size 10 x 20 x 5 mm, geometry from box.sld
        - object Box at (696768, 103.35, 13.17) mm, rotated rx -0.49 ry 0.34 rz 17 deg, size 10 x 20 x 5 mm, geometry from box.sld
        - object Box at (696167, 103.35, 13.17) mm, rotated rx -0.27 ry 0.53 rz 44.9 deg, size 10 x 20 x 5 mm, geometry from box.sld
        - object Box at (695554, 103.35, 13.17) mm, rotated rx -0.37 ry 0.46 rz 33.31 deg, size 10 x 20 x 5 mm, geometry from box.sld
        - object Box at (694953, 103.35, 13.17) mm, rotated rx -0.59 ry -0.04 rz -22.04 deg, size 10 x 20 x 5 mm, geometry from box.sld
        - object Box at (694333, 103.35, 13.17) mm, rotated rx -0.53 ry 0.27 rz 9.42 deg, size 10 x 20 x 5 mm, geometry from box.sld
        - object Box at (693726, 103.35, 13.17) mm, rotated rx -0.58 ry -0.15 rz -32.46 deg, size 10 x 20 x 5 mm, geometry from box.sld
        - object Box at (693129, 103.35, 13.17) mm, rotated rx -0.57 ry -0.16 rz -34.07 deg, size 10 x 20 x 5 mm, geometry from box.sld
        - object Box at (692511, 103.35, 13.17) mm, rotated rx -0.46 ry 0.37 rz 20.63 deg, size 10 x 20 x 5 mm, geometry from box.sld
        - object Box at (691916, 103.35, 13.17) mm, rotated rx -0.53 ry -0.26 rz -43.89 deg, size 10 x 20 x 5 mm, geometry from box.sld
        - object Box at (691310, 103.35, 13.17) mm, rotated rx -0.37 ry 0.46 rz 33.32 deg, size 10 x 20 x 5 mm, geometry from box.sld
        - object Box at (690702, 103.35, 13.17) mm, rotated rx -0.58 ry -0.12 rz -29.89 deg, size 10 x 20 x 5 mm, geometry from box.sld
        - object Box at (690083, 103.35, 13.17) mm, rotated rx -0.57 ry 0.16 rz -2.2 deg, size 10 x 20 x 5 mm, geometry from box.sld
        - object Box at (689452, 103.35, 13.17) mm, rotated rx -0.59 ry 0.05 rz -13.09 deg, size 10 x 20 x 5 mm, geometry from box.sld
        - object Box at (688852, 103.35, 13.17) mm, rotated rx -0.39 ry 0.45 rz 30.45 deg, size 10 x 20 x 5 mm, geometry from box.sld
        - object Box at (688240, 103.35, 13.17) mm, rotated rx -0.42 ry 0.42 rz 26.77 deg, size 10 x 20 x 5 mm, geometry from box.sld
        - object Box at (687617, 103.35, 13.17) mm, rotated rx -0.59 ry -0.1 rz -27.42 deg, size 10 x 20 x 5 mm, geometry from box.sld
        - object Box at (686998, 103.35, 13.17) mm, rotated rx -0.47 ry 0.37 rz 20.14 deg, size 10 x 20 x 5 mm, geometry from box.sld
        - object Box at (686383, 103.35, 13.17) mm, rotated rx -0.41 ry 0.43 rz 28.79 deg, size 10 x 20 x 5 mm, geometry from box.sld
        - object Box at (685759, 103.35, 13.17) mm, rotated rx -0.57 ry -0.18 rz -35.37 deg, size 10 x 20 x 5 mm, geometry from box.sld
        - object Box at (685124, 103.35, 13.17) mm, rotated rx -0.41 ry 0.43 rz 28.79 deg, size 10 x 20 x 5 mm, geometry from box.sld
        - object Box at (684514, 103.35, 13.17) mm, rotated rx -0.45 ry 0.39 rz 23.21 deg, size 10 x 20 x 5 mm, geometry from box.sld
        - object Box at (683902, 103.35, 13.17) mm, rotated rx -0.28 ry 0.52 rz 43.82 deg, size 10 x 20 x 5 mm, geometry from box.sld
        - object Box at (683303, 103.35, 13.17) mm, rotated rx -0.4 ry 0.43 rz 28.84 deg, size 10 x 20 x 5 mm, geometry from box.sld
        - object Box at (682690, 103.35, 13.17) mm, rotated rx -0.51 ry 0.3 rz 12.46 deg, size 10 x 20 x 5 mm, geometry from box.sld
        - object Box at (682071, 103.35, 13.17) mm, rotated rx -0.58 ry 0.14 rz -4.32 deg, size 10 x 20 x 5 mm, geometry from box.sld
        - object Box at (681452, 103.35, 13.17) mm, rotated rx -0.59 ry 0.07 rz -11.71 deg, size 10 x 20 x 5 mm, geometry from box.sld
        - object Box at (680819, 103.35, 13.17) mm, rotated rx -0.58 ry 0.11 rz -7.05 deg, size 10 x 20 x 5 mm, geometry from box.sld
        - object Box at (680187, 103.35, 13.17) mm, rotated rx -0.43 ry 0.4 rz 24.78 deg, size 10 x 20 x 5 mm, geometry from box.sld
        - object Box at (679572, 103.35, 13.17) mm, rotated rx -0.44 ry 0.4 rz 24.26 deg, size 10 x 20 x 5 mm, geometry from box.sld
        - object Box at (678984, 103.35, 13.17) mm, rotated rx -0.58 ry 0.15 rz -3.98 deg, size 10 x 20 x 5 mm, geometry from box.sld
        - object Box at (678382, 103.35, 13.17) mm, rotated rx -0.35 ry 0.48 rz 35.28 deg, size 10 x 20 x 5 mm, geometry from box.sld
        - object Box at (677789, 103.35, 13.17) mm, rotated rx -0.57 ry -0.17 rz -35.2 deg, size 10 x 20 x 5 mm, geometry from box.sld
        - object Box at (677203, 103.35, 13.17) mm, rotated rx -0.48 ry 0.35 rz 18.23 deg, size 10 x 20 x 5 mm, geometry from box.sld
        - object Box at (676608, 103.35, 13.17) mm, rotated rx -0.59 ry 0.03 rz -14.98 deg, size 10 x 20 x 5 mm, geometry from box.sld
        - object Box at (676012, 103.35, 13.17) mm, rotated rx -0.41 ry 0.43 rz 28.4 deg, size 10 x 20 x 5 mm, geometry from box.sld
        - object Box at (675418, 103.35, 13.17) mm, rotated rx -0.5 ry 0.31 rz 13.8 deg, size 10 x 20 x 5 mm, geometry from box.sld
        - object Box at (674814, 103.35, 13.17) mm, rotated rx -0.59 ry 0.08 rz -10.17 deg, size 10 x 20 x 5 mm, geometry from box.sld
        - object Box at (674215, 103.35, 13.17) mm, rotated rx -0.58 ry 0.13 rz -5.17 deg, size 10 x 20 x 5 mm, geometry from box.sld
        - object Box at (673617, 103.35, 13.17) mm, rotated rx -0.4 ry 0.44 rz 29.04 deg, size 10 x 20 x 5 mm, geometry from box.sld
        - object Box at (673020, 103.35, 13.17) mm, rotated rx -0.47 ry 0.36 rz 18.88 deg, size 10 x 20 x 5 mm, geometry from box.sld
        - object Box at (672417, 103.35, 13.17) mm, rotated rx -0.35 ry 0.48 rz 35.99 deg, size 10 x 20 x 5 mm, geometry from box.sld
        - object Box at (671818, 103.35, 13.17) mm, rotated rx -0.59 ry -0.07 rz -24.76 deg, size 10 x 20 x 5 mm, geometry from box.sld
        - object Box at (671218, 103.35, 13.17) mm, rotated rx -0.56 ry 0.2 rz 1.65 deg, size 10 x 20 x 5 mm, geometry from box.sld
        - object Box at (670618, 103.35, 13.17) mm, rotated rx -0.59 ry -0.03 rz -20.92 deg, size 10 x 20 x 5 mm, geometry from box.sld
        - object Box at (670023, 103.35, 13.17) mm, rotated rx -0.57 ry -0.18 rz -35.6 deg, size 10 x 20 x 5 mm, geometry from box.sld
        - object Box at (669422, 103.35, 13.17) mm, rotated rx -0.41 ry 0.43 rz 28.58 deg, size 10 x 20 x 5 mm, geometry from box.sld
        - object Box at (668822, 103.35, 13.17) mm, rotated rx -0.3 ry 0.51 rz 41.32 deg, size 10 x 20 x 5 mm, geometry from box.sld
        - object Box at (668225, 103.35, 13.17) mm, rotated rx -0.45 ry 0.39 rz 23.15 deg, size 10 x 20 x 5 mm, geometry from box.sld
        - object Box at (667626, 103.35, 13.17) mm, rotated rx -0.46 ry 0.38 rz 21.46 deg, size 10 x 20 x 5 mm, geometry from box.sld
        - object Box at (667027, 103.35, 13.17) mm, rotated rx -0.29 ry 0.52 rz 42.9 deg, size 10 x 20 x 5 mm, geometry from box.sld
        - object Box at (666421, 103.35, 13.17) mm, rotated rx -0.59 ry 0.06 rz -12.81 deg, size 10 x 20 x 5 mm, geometry from box.sld
        - object Box at (665822, 103.35, 13.17) mm, rotated rx -0.51 ry 0.3 rz 11.78 deg, size 10 x 20 x 5 mm, geometry from box.sld
        - object Box at (665216, 103.35, 13.17) mm, rotated rx -0.37 ry 0.47 rz 33.45 deg, size 10 x 20 x 5 mm, geometry from box.sld
        - object Box at (664615, 103.35, 13.17) mm, rotated rx -0.59 ry -0.01 rz -19.28 deg, size 10 x 20 x 5 mm, geometry from box.sld
        - object Box at (664014, 103.35, 13.17) mm, rotated rx -0.49 ry 0.33 rz 15.82 deg, size 10 x 20 x 5 mm, geometry from box.sld
        - object Box at (663411, 103.35, 13.17) mm, rotated rx -0.54 ry 0.25 rz 6.26 deg, size 10 x 20 x 5 mm, geometry from box.sld
        - object Box at (662813, 103.35, 13.17) mm, rotated rx -0.59 ry -0.07 rz -25.25 deg, size 10 x 20 x 5 mm, geometry from box.sld
        - object Box at (662207, 103.35, 13.17) mm, rotated rx -0.47 ry 0.36 rz 18.9 deg, size 10 x 20 x 5 mm, geometry from box.sld
        - object Box at (661609, 103.35, 13.17) mm, rotated rx -0.57 ry 0.16 rz -2.74 deg, size 10 x 20 x 5 mm, geometry from box.sld
        - object Box at (661009, 103.35, 13.17) mm, rotated rx -0.58 ry -0.13 rz -30.45 deg, size 10 x 20 x 5 mm, geometry from box.sld
        - object Box at (660406, 103.35, 13.17) mm, rotated rx -0.55 ry 0.23 rz 4.34 deg, size 10 x 20 x 5 mm, geometry from box.sld
        - object Box at (659802, 103.35, 13.17) mm, rotated rx -0.54 ry 0.25 rz 6.84 deg, size 10 x 20 x 5 mm, geometry from box.sld
        - object Box at (659198, 103.35, 13.17) mm, rotated rx -0.41 ry 0.43 rz 28.48 deg, size 10 x 20 x 5 mm, geometry from box.sld
        - object Box at (658593, 103.35, 13.17) mm, rotated rx -0.54 ry 0.24 rz 5.92 deg, size 10 x 20 x 5 mm, geometry from box.sld
        - object Box at (657989, 103.35, 13.17) mm, rotated rx -0.56 ry 0.21 rz 2.35 deg, size 10 x 20 x 5 mm, geometry from box.sld
        - object Box at (657382, 103.35, 13.17) mm, rotated rx -0.59 ry 0.06 rz -12.69 deg, size 10 x 20 x 5 mm, geometry from box.sld
        - object Box at (656774, 103.35, 13.17) mm, rotated rx -0.55 ry 0.22 rz 3.69 deg, size 10 x 20 x 5 mm, geometry from box.sld
        - object Box at (656171, 103.35, 13.17) mm, rotated rx -0.42 ry 0.42 rz 27.15 deg, size 10 x 20 x 5 mm, geometry from box.sld
        - object Box at (655567, 103.35, 13.17) mm, rotated rx -0.56 ry -0.2 rz -37.52 deg, size 10 x 20 x 5 mm, geometry from box.sld
        - object Box at (654959, 103.35, 13.17) mm, rotated rx -0.57 ry -0.18 rz -36.01 deg, size 10 x 20 x 5 mm, geometry from box.sld
        - object Box at (654352, 103.35, 13.17) mm, rotated rx -0.58 ry -0.14 rz -31.93 deg, size 10 x 20 x 5 mm, geometry from box.sld
        - object Box at (653741, 103.35, 13.17) mm, rotated rx -0.56 ry -0.2 rz -37.76 deg, size 10 x 20 x 5 mm, geometry from box.sld
        - object Box at (653117, 103.35, 13.17) mm, rotated rx -0.58 ry 0.14 rz -4.41 deg, size 10 x 20 x 5 mm, geometry from box.sld
        - object Box at (652513, 103.35, 13.17) mm, rotated rx -0.39 ry 0.45 rz 31.18 deg, size 10 x 20 x 5 mm, geometry from box.sld
        - object Box at (651905, 103.35, 13.17) mm, rotated rx -0.59 ry 0.09 rz -8.99 deg, size 10 x 20 x 5 mm, geometry from box.sld
        - object Box at (651292, 103.35, 13.17) mm, rotated rx -0.39 ry 0.45 rz 31.01 deg, size 10 x 20 x 5 mm, geometry from box.sld
        - object Box at (650684, 103.35, 13.17) mm, rotated rx -0.58 ry -0.14 rz -31.69 deg, size 10 x 20 x 5 mm, geometry from box.sld
        - object Box at (650061, 103.35, 13.17) mm, rotated rx -0.55 ry 0.23 rz 4.83 deg, size 10 x 20 x 5 mm, geometry from box.sld
        - object Box at (649447, 103.35, 13.17) mm, rotated rx -0.51 ry 0.31 rz 12.97 deg, size 10 x 20 x 5 mm, geometry from box.sld
        - object Box at (648835, 103.35, 13.17) mm, rotated rx -0.52 ry 0.29 rz 11.46 deg, size 10 x 20 x 5 mm, geometry from box.sld
        - object Box at (648218, 103.35, 13.17) mm, rotated rx -0.58 ry -0.11 rz -28.4 deg, size 10 x 20 x 5 mm, geometry from box.sld
        - object Box at (647607, 103.35, 13.17) mm, rotated rx -0.56 ry 0.19 rz 0.07 deg, size 10 x 20 x 5 mm, geometry from box.sld
        - object Box at (646995, 103.35, 13.17) mm, rotated rx -0.57 ry 0.17 rz -1.68 deg, size 10 x 20 x 5 mm, geometry from box.sld
        - object Box at (646378, 103.35, 13.17) mm, rotated rx -0.59 ry 0.04 rz -14 deg, size 10 x 20 x 5 mm, geometry from box.sld
        - object Box at (645763, 103.35, 13.17) mm, rotated rx -0.42 ry 0.42 rz 26.45 deg, size 10 x 20 x 5 mm, geometry from box.sld
        - object Box at (645143, 103.35, 13.17) mm, rotated rx -0.45 ry 0.39 rz 23.01 deg, size 10 x 20 x 5 mm, geometry from box.sld
        - object Box at (644523, 103.35, 13.17) mm, rotated rx -0.45 ry 0.38 rz 21.86 deg, size 10 x 20 x 5 mm, geometry from box.sld
        - object Box at (643906, 103.35, 13.17) mm, rotated rx -0.54 ry 0.25 rz 6.22 deg, size 10 x 20 x 5 mm, geometry from box.sld
        - object Box at (643287, 103.35, 13.17) mm, rotated rx -0.56 ry 0.21 rz 2.5 deg, size 10 x 20 x 5 mm, geometry from box.sld
        - object Box at (642673, 103.35, 13.17) mm, rotated rx -0.56 ry 0.2 rz 1.34 deg, size 10 x 20 x 5 mm, geometry from box.sld
        - object Box at (642052, 103.35, 13.17) mm, rotated rx -0.58 ry -0.12 rz -30.09 deg, size 10 x 20 x 5 mm, geometry from box.sld
        - object Box at (641435, 103.35, 13.17) mm, rotated rx -0.59 ry 0 rz -18.57 deg, size 10 x 20 x 5 mm, geometry from box.sld
        - object Box at (640822, 103.35, 13.17) mm, rotated rx -0.3 ry 0.51 rz 41.89 deg, size 10 x 20 x 5 mm, geometry from box.sld
        - object Box at (640200, 103.35, 13.17) mm, rotated rx -0.58 ry -0.13 rz -30.52 deg, size 10 x 20 x 5 mm, geometry from box.sld
        - object Box at (639583, 103.35, 13.17) mm, rotated rx -0.59 ry -0.05 rz -23.07 deg, size 10 x 20 x 5 mm, geometry from box.sld
        - object Box at (638963, 103.35, 13.17) mm, rotated rx -0.58 ry 0.12 rz -6.56 deg, size 10 x 20 x 5 mm, geometry from box.sld
        - object Box at (638350, 103.35, 13.17) mm, rotated rx -0.55 ry -0.21 rz -39.39 deg, size 10 x 20 x 5 mm, geometry from box.sld
        - object Box at (637726, 103.35, 13.17) mm, rotated rx -0.59 ry 0.05 rz -13.32 deg, size 10 x 20 x 5 mm, geometry from box.sld
        - object Box at (637103, 103.35, 13.17) mm, rotated rx -0.28 ry 0.53 rz 44.04 deg, size 10 x 20 x 5 mm, geometry from box.sld
        - object Box at (636484, 103.35, 13.17) mm, rotated rx -0.59 ry 0.06 rz -12.15 deg, size 10 x 20 x 5 mm, geometry from box.sld
        - object Box at (635864, 103.35, 13.17) mm, rotated rx -0.44 ry 0.39 rz 23.39 deg, size 10 x 20 x 5 mm, geometry from box.sld
        - object Box at (635248, 103.35, 13.17) mm, rotated rx -0.5 ry 0.32 rz 13.92 deg, size 10 x 20 x 5 mm, geometry from box.sld
        - object Box at (634626, 103.35, 13.17) mm, rotated rx -0.59 ry 0 rz -18.19 deg, size 10 x 20 x 5 mm, geometry from box.sld
        - object Box at (634006, 103.35, 13.17) mm, rotated rx -0.56 ry -0.2 rz -37.64 deg, size 10 x 20 x 5 mm, geometry from box.sld
        - object Box at (633383, 103.35, 13.17) mm, rotated rx -0.58 ry 0.12 rz -6.51 deg, size 10 x 20 x 5 mm, geometry from box.sld
        - object Box at (632760, 103.35, 13.17) mm, rotated rx -0.59 ry -0.03 rz -20.64 deg, size 10 x 20 x 5 mm, geometry from box.sld
        - object Box at (632132, 103.35, 13.17) mm, rotated rx -0.57 ry -0.17 rz -35.21 deg, size 10 x 20 x 5 mm, geometry from box.sld
        - object Box at (631510, 103.35, 13.17) mm, rotated rx -0.54 ry 0.24 rz 5.49 deg, size 10 x 20 x 5 mm, geometry from box.sld
        - object Box at (630887, 103.35, 13.17) mm, rotated rx -0.55 ry 0.23 rz 4.57 deg, size 10 x 20 x 5 mm, geometry from box.sld
        - object Box at (630262, 103.35, 13.17) mm, rotated rx -0.59 ry -0.05 rz -22.54 deg, size 10 x 20 x 5 mm, geometry from box.sld
        - object Box at (629638, 103.35, 13.17) mm, rotated rx -0.58 ry 0.14 rz -4.7 deg, size 10 x 20 x 5 mm, geometry from box.sld
        - object Box at (629010, 103.35, 13.17) mm, rotated rx -0.29 ry 0.52 rz 43 deg, size 10 x 20 x 5 mm, geometry from box.sld
        - object Box at (628378, 103.35, 13.17) mm, rotated rx -0.4 ry 0.44 rz 29.16 deg, size 10 x 20 x 5 mm, geometry from box.sld
        - object Box at (627744, 103.35, 13.17) mm, rotated rx -0.57 ry -0.16 rz -33.99 deg, size 10 x 20 x 5 mm, geometry from box.sld
        - object Box at (627118, 103.35, 13.17) mm, rotated rx -0.49 ry 0.34 rz 16.3 deg, size 10 x 20 x 5 mm, geometry from box.sld
        - object Box at (626495, 103.35, 13.17) mm, rotated rx -0.59 ry 0.01 rz -17.32 deg, size 10 x 20 x 5 mm, geometry from box.sld
        - object Box at (625863, 103.35, 13.17) mm, rotated rx -0.52 ry 0.29 rz 10.77 deg, size 10 x 20 x 5 mm, geometry from box.sld
        - object Box at (625243, 103.35, 13.17) mm, rotated rx -0.57 ry -0.17 rz -34.49 deg, size 10 x 20 x 5 mm, geometry from box.sld
        - object Box at (624615, 103.35, 13.17) mm, rotated rx -0.58 ry -0.14 rz -32.16 deg, size 10 x 20 x 5 mm, geometry from box.sld
        - object Box at (623993, 103.35, 13.17) mm, rotated rx -0.58 ry 0.12 rz -6.22 deg, size 10 x 20 x 5 mm, geometry from box.sld
        - object Box at (623362, 103.35, 13.17) mm, rotated rx -0.58 ry -0.13 rz -30.55 deg, size 10 x 20 x 5 mm, geometry from box.sld
        - object Box at (622730, 103.35, 13.17) mm, rotated rx -0.59 ry 0.04 rz -13.91 deg, size 10 x 20 x 5 mm, geometry from box.sld
        - object Box at (622100, 103.35, 13.17) mm, rotated rx -0.54 ry -0.24 rz -41.52 deg, size 10 x 20 x 5 mm, geometry from box.sld
        - object Box at (621468, 103.35, 13.17) mm, rotated rx -0.59 ry 0.04 rz -13.83 deg, size 10 x 20 x 5 mm, geometry from box.sld
        - object Box at (620839, 103.35, 13.17) mm, rotated rx -0.59 ry 0.07 rz -11.48 deg, size 10 x 20 x 5 mm, geometry from box.sld
        - object Box at (620215, 103.35, 13.17) mm, rotated rx -0.56 ry -0.21 rz -38.38 deg, size 10 x 20 x 5 mm, geometry from box.sld
        - object Box at (619580, 103.35, 13.17) mm, rotated rx -0.54 ry -0.24 rz -41.69 deg, size 10 x 20 x 5 mm, geometry from box.sld
        - object Box at (618943, 103.35, 13.17) mm, rotated rx -0.59 ry -0.03 rz -20.9 deg, size 10 x 20 x 5 mm, geometry from box.sld
        - object Box at (618309, 103.35, 13.17) mm, rotated rx -0.59 ry 0.02 rz -16.03 deg, size 10 x 20 x 5 mm, geometry from box.sld
        - object Box at (617676, 103.35, 13.17) mm, rotated rx -0.57 ry 0.17 rz -1.14 deg, size 10 x 20 x 5 mm, geometry from box.sld
        - object Box at (617047, 103.35, 13.17) mm, rotated rx -0.53 ry -0.26 rz -44.62 deg, size 10 x 20 x 5 mm, geometry from box.sld
        - object Box at (616407, 103.35, 13.17) mm, rotated rx -0.42 ry 0.42 rz 27.41 deg, size 10 x 20 x 5 mm, geometry from box.sld
        - object Box at (615775, 103.35, 13.17) mm, rotated rx -0.53 ry 0.27 rz 9.19 deg, size 10 x 20 x 5 mm, geometry from box.sld
        - object Box at (615115, 103.35, 13.17) mm, rotated rx -0.57 ry -0.16 rz -33.76 deg, size 10 x 20 x 5 mm, geometry from box.sld
        - object Box at (614483, 103.35, 13.17) mm, rotated rx -0.59 ry -0.01 rz -18.74 deg, size 10 x 20 x 5 mm, geometry from box.sld
        - object Box at (613850, 103.35, 13.17) mm, rotated rx -0.59 ry 0.1 rz -8.92 deg, size 10 x 20 x 5 mm, geometry from box.sld
        - object Box at (613210, 103.35, 13.17) mm, rotated rx -0.59 ry 0.07 rz -11.25 deg, size 10 x 20 x 5 mm, geometry from box.sld
        - object Box at (612577, 103.35, 13.17) mm, rotated rx -0.48 ry 0.35 rz 18.15 deg, size 10 x 20 x 5 mm, geometry from box.sld
        - object Box at (611939, 103.35, 13.17) mm, rotated rx -0.58 ry 0.12 rz -6.97 deg, size 10 x 20 x 5 mm, geometry from box.sld
        - object Box at (611304, 103.35, 13.17) mm, rotated rx -0.54 ry -0.24 rz -41.87 deg, size 10 x 20 x 5 mm, geometry from box.sld
        - object Box at (610659, 103.35, 13.17) mm, rotated rx -0.35 ry 0.48 rz 35.34 deg, size 10 x 20 x 5 mm, geometry from box.sld
        - object Box at (610027, 103.35, 13.17) mm, rotated rx -0.48 ry 0.35 rz 18.01 deg, size 10 x 20 x 5 mm, geometry from box.sld
        - object Box at (609383, 103.35, 13.17) mm, rotated rx -0.56 ry 0.21 rz 2.12 deg, size 10 x 20 x 5 mm, geometry from box.sld
        - object Box at (608747, 103.35, 13.17) mm, rotated rx -0.58 ry -0.12 rz -29.43 deg, size 10 x 20 x 5 mm, geometry from box.sld
        - object Box at (607940, 103.35, 13.17) mm, rotated rx -0.46 ry 0.37 rz 20.3 deg, size 10 x 20 x 5 mm, geometry from box.sld
        - object Box at (607304, 103.35, 13.17) mm, rotated rx -0.44 ry 0.4 rz 23.67 deg, size 10 x 20 x 5 mm, geometry from box.sld
        - object Box at (606667, 103.35, 13.17) mm, rotated rx -0.49 ry 0.34 rz 16.78 deg, size 10 x 20 x 5 mm, geometry from box.sld
        - object Box at (606022, 103.35, 13.17) mm, rotated rx -0.59 ry 0.07 rz -11.33 deg, size 10 x 20 x 5 mm, geometry from box.sld
        - object Box at (605376, 103.35, 13.17) mm, rotated rx -0.59 ry 0.02 rz -16.55 deg, size 10 x 20 x 5 mm, geometry from box.sld
        - object Box at (604734, 103.35, 13.17) mm, rotated rx -0.59 ry 0.1 rz -8.66 deg, size 10 x 20 x 5 mm, geometry from box.sld
        - object Box at (604092, 103.35, 13.17) mm, rotated rx -0.58 ry -0.14 rz -32.07 deg, size 10 x 20 x 5 mm, geometry from box.sld
        - object Box at (603453, 103.35, 13.17) mm, rotated rx -0.59 ry 0.09 rz -9.58 deg, size 10 x 20 x 5 mm, geometry from box.sld
        - object Box at (602812, 103.35, 13.17) mm, rotated rx -0.5 ry 0.32 rz 15.02 deg, size 10 x 20 x 5 mm, geometry from box.sld
        - object Box at (602165, 103.35, 13.17) mm, rotated rx -0.54 ry -0.24 rz -42 deg, size 10 x 20 x 5 mm, geometry from box.sld
        - object Box at (601520, 103.35, 13.17) mm, rotated rx -0.29 ry 0.52 rz 42.23 deg, size 10 x 20 x 5 mm, geometry from box.sld
        - object Box at (600809, 103.35, 13.17) mm, rotated rx -0.59 ry -0.01 rz -19.36 deg, size 10 x 20 x 5 mm, geometry from box.sld
        - object Box at (600167, 103.35, 13.17) mm, rotated rx -0.58 ry 0.15 rz -4 deg, size 10 x 20 x 5 mm, geometry from box.sld
        - object Box at (599795, 103.35, 13.17) mm, rotated rx -0.54 ry 0.25 rz 7.2 deg, size 10 x 20 x 5 mm, geometry from box.sld
        - object Box at (599156, 103.35, 13.17) mm, rotated rx -0.34 ry 0.49 rz 37.18 deg, size 10 x 20 x 5 mm, geometry from box.sld
        - object Box at (598514, 103.35, 13.17) mm, rotated rx -0.59 ry -0.01 rz -19.42 deg, size 10 x 20 x 5 mm, geometry from box.sld
        - object Box at (597869, 103.35, 13.17) mm, rotated rx -0.41 ry 0.43 rz 27.83 deg, size 10 x 20 x 5 mm, geometry from box.sld
        - object Box at (597212, 103.35, 13.17) mm, rotated rx -0.28 ry 0.53 rz 44.09 deg, size 10 x 20 x 5 mm, geometry from box.sld
        - object Box at (596568, 103.35, 13.17) mm, rotated rx -0.58 ry -0.12 rz -30.05 deg, size 10 x 20 x 5 mm, geometry from box.sld
        - object Box at (595924, 103.35, 13.17) mm, rotated rx -0.32 ry 0.5 rz 38.72 deg, size 10 x 20 x 5 mm, geometry from box.sld
        - object Box at (595280, 103.35, 13.17) mm, rotated rx -0.59 ry 0.07 rz -11.2 deg, size 10 x 20 x 5 mm, geometry from box.sld
        - object Box at (594637, 103.35, 13.17) mm, rotated rx -0.38 ry 0.46 rz 32.34 deg, size 10 x 20 x 5 mm, geometry from box.sld
        - object Box at (593993, 103.35, 13.17) mm, rotated rx -0.43 ry 0.41 rz 25.55 deg, size 10 x 20 x 5 mm, geometry from box.sld
        - object Box at (593344, 103.35, 13.17) mm, rotated rx -0.36 ry 0.47 rz 33.95 deg, size 10 x 20 x 5 mm, geometry from box.sld
        - object Box at (592697, 103.35, 13.17) mm, rotated rx -0.59 ry 0.03 rz -14.91 deg, size 10 x 20 x 5 mm, geometry from box.sld
        - object Box at (592050, 103.35, 13.17) mm, rotated rx -0.58 ry 0.11 rz -7.21 deg, size 10 x 20 x 5 mm, geometry from box.sld
        - object Box at (591404, 103.35, 13.17) mm, rotated rx -0.59 ry 0 rz -17.72 deg, size 10 x 20 x 5 mm, geometry from box.sld
        - object Box at (590752, 103.35, 13.17) mm, rotated rx -0.59 ry -0.04 rz -22.18 deg, size 10 x 20 x 5 mm, geometry from box.sld
        - object Box at (590097, 103.35, 13.17) mm, rotated rx -0.41 ry 0.43 rz 27.88 deg, size 10 x 20 x 5 mm, geometry from box.sld
        - object Box at (589451, 103.35, 13.17) mm, rotated rx -0.38 ry 0.45 rz 31.65 deg, size 10 x 20 x 5 mm, geometry from box.sld
        - object Box at (588800, 103.35, 13.17) mm, rotated rx -0.57 ry 0.16 rz -2.89 deg, size 10 x 20 x 5 mm, geometry from box.sld
        - object Box at (588151, 103.35, 13.17) mm, rotated rx -0.51 ry 0.31 rz 13.06 deg, size 10 x 20 x 5 mm, geometry from box.sld
        - object Box at (587500, 103.35, 13.17) mm, rotated rx -0.41 ry 0.43 rz 28.5 deg, size 10 x 20 x 5 mm, geometry from box.sld
        - object Box at (586850, 103.35, 13.17) mm, rotated rx -0.54 ry 0.24 rz 5.73 deg, size 10 x 20 x 5 mm, geometry from box.sld
        - object Box at (586202, 103.35, 13.17) mm, rotated rx -0.33 ry 0.49 rz 37.8 deg, size 10 x 20 x 5 mm, geometry from box.sld
        - object Box at (585554, 103.35, 13.17) mm, rotated rx -0.59 ry 0.07 rz -11.77 deg, size 10 x 20 x 5 mm, geometry from box.sld
        - object Box at (584899, 103.35, 13.17) mm, rotated rx -0.46 ry 0.38 rz 21.78 deg, size 10 x 20 x 5 mm, geometry from box.sld
        - object Box at (584245, 103.35, 13.17) mm, rotated rx -0.3 ry 0.51 rz 41.26 deg, size 10 x 20 x 5 mm, geometry from box.sld
        - object Box at (583589, 103.35, 13.17) mm, rotated rx -0.56 ry 0.2 rz 1.88 deg, size 10 x 20 x 5 mm, geometry from box.sld
        - object Box at (582911, 103.35, 13.17) mm, rotated rx -0.57 ry -0.17 rz -34.78 deg, size 10 x 20 x 5 mm, geometry from box.sld
        - object Box at (582260, 103.35, 13.17) mm, rotated rx -0.54 ry 0.25 rz 6.45 deg, size 10 x 20 x 5 mm, geometry from box.sld
        - object Box at (581605, 103.35, 13.17) mm, rotated rx -0.58 ry -0.1 rz -28.1 deg, size 10 x 20 x 5 mm, geometry from box.sld
        - object Box at (580954, 103.35, 13.17) mm, rotated rx -0.59 ry -0.05 rz -23.05 deg, size 10 x 20 x 5 mm, geometry from box.sld
        - object Box at (580302, 103.35, 13.17) mm, rotated rx -0.39 ry 0.45 rz 30.98 deg, size 10 x 20 x 5 mm, geometry from box.sld
        - object Box at (579646, 103.35, 13.17) mm, rotated rx -0.37 ry 0.47 rz 33.82 deg, size 10 x 20 x 5 mm, geometry from box.sld
        - object Box at (578995, 103.35, 13.17) mm, rotated rx -0.35 ry 0.48 rz 35.46 deg, size 10 x 20 x 5 mm, geometry from box.sld
        - object Box at (578339, 103.35, 13.17) mm, rotated rx -0.53 ry 0.26 rz 7.57 deg, size 10 x 20 x 5 mm, geometry from box.sld
        - object Box at (577681, 103.35, 13.17) mm, rotated rx -0.59 ry 0.04 rz -14.04 deg, size 10 x 20 x 5 mm, geometry from box.sld
        - object Box at (577021, 103.35, 13.17) mm, rotated rx -0.57 ry 0.16 rz -2.08 deg, size 10 x 20 x 5 mm, geometry from box.sld
        - object Box at (576365, 103.35, 13.17) mm, rotated rx -0.31 ry 0.51 rz 40.7 deg, size 10 x 20 x 5 mm, geometry from box.sld
        - object Box at (575709, 103.35, 13.17) mm, rotated rx -0.59 ry 0.06 rz -12.05 deg, size 10 x 20 x 5 mm, geometry from box.sld
        - object Box at (575053, 103.35, 13.17) mm, rotated rx -0.52 ry 0.28 rz 10.37 deg, size 10 x 20 x 5 mm, geometry from box.sld
        - object Box at (574394, 103.35, 13.17) mm, rotated rx -0.35 ry 0.48 rz 35.57 deg, size 10 x 20 x 5 mm, geometry from box.sld
        - object Box at (573729, 103.35, 13.17) mm, rotated rx -0.44 ry 0.4 rz 24.08 deg, size 10 x 20 x 5 mm, geometry from box.sld
        - object Box at (573074, 103.35, 13.17) mm, rotated rx -0.59 ry 0.03 rz -15.05 deg, size 10 x 20 x 5 mm, geometry from box.sld
        - object Box at (572413, 103.35, 13.17) mm, rotated rx -0.5 ry 0.32 rz 14.01 deg, size 10 x 20 x 5 mm, geometry from box.sld
        - object Box at (571748, 103.35, 13.17) mm, rotated rx -0.27 ry 0.53 rz 44.57 deg, size 10 x 20 x 5 mm, geometry from box.sld
        - object Box at (571092, 103.35, 13.17) mm, rotated rx -0.57 ry -0.16 rz -33.33 deg, size 10 x 20 x 5 mm, geometry from box.sld
        - object Box at (570436, 103.35, 13.17) mm, rotated rx -0.37 ry 0.47 rz 33.82 deg, size 10 x 20 x 5 mm, geometry from box.sld
        - object Box at (569774, 103.35, 13.17) mm, rotated rx -0.53 ry -0.26 rz -44.07 deg, size 10 x 20 x 5 mm, geometry from box.sld
        - object Box at (569112, 103.35, 13.17) mm, rotated rx -0.45 ry 0.39 rz 23.22 deg, size 10 x 20 x 5 mm, geometry from box.sld
        - object Box at (568448, 103.35, 13.17) mm, rotated rx -0.5 ry 0.32 rz 14.54 deg, size 10 x 20 x 5 mm, geometry from box.sld
        - object Box at (567790, 103.35, 13.17) mm, rotated rx -0.5 ry 0.32 rz 14.6 deg, size 10 x 20 x 5 mm, geometry from box.sld
        - object Box at (567128, 103.35, 13.17) mm, rotated rx -0.47 ry 0.37 rz 19.99 deg, size 10 x 20 x 5 mm, geometry from box.sld
        - object Box at (566463, 103.35, 13.17) mm, rotated rx -0.58 ry -0.15 rz -32.39 deg, size 10 x 20 x 5 mm, geometry from box.sld
        - object Box at (565803, 103.35, 13.17) mm, rotated rx -0.51 ry 0.3 rz 12.46 deg, size 10 x 20 x 5 mm, geometry from box.sld
        - object Box at (565143, 103.35, 13.17) mm, rotated rx -0.52 ry 0.29 rz 11.08 deg, size 10 x 20 x 5 mm, geometry from box.sld
        - object Box at (564479, 103.35, 13.17) mm, rotated rx -0.54 ry 0.25 rz 6.31 deg, size 10 x 20 x 5 mm, geometry from box.sld
        - object Box at (563813, 103.35, 13.17) mm, rotated rx -0.29 ry 0.52 rz 43.13 deg, size 10 x 20 x 5 mm, geometry from box.sld
        - object Box at (563148, 103.35, 13.17) mm, rotated rx -0.43 ry 0.41 rz 25.42 deg, size 10 x 20 x 5 mm, geometry from box.sld
        - object Box at (562485, 103.35, 13.17) mm, rotated rx -0.57 ry 0.15 rz -3.19 deg, size 10 x 20 x 5 mm, geometry from box.sld
        - object Box at (561822, 103.35, 13.17) mm, rotated rx -0.56 ry 0.18 rz -0.29 deg, size 10 x 20 x 5 mm, geometry from box.sld
        - object Box at (561158, 103.35, 13.17) mm, rotated rx -0.5 ry 0.33 rz 15.07 deg, size 10 x 20 x 5 mm, geometry from box.sld
        - object Box at (560485, 103.35, 13.17) mm, rotated rx -0.54 ry -0.24 rz -42.13 deg, size 10 x 20 x 5 mm, geometry from box.sld
        - object Box at (559815, 103.35, 13.17) mm, rotated rx -0.52 ry 0.28 rz 10.14 deg, size 10 x 20 x 5 mm, geometry from box.sld
        - object Box at (559156, 103.35, 13.17) mm, rotated rx -0.59 ry 0.01 rz -17 deg, size 10 x 20 x 5 mm, geometry from box.sld
        - object Box at (558492, 103.35, 13.17) mm, rotated rx -0.29 ry 0.52 rz 43.04 deg, size 10 x 20 x 5 mm, geometry from box.sld
        - object Box at (557824, 103.35, 13.17) mm, rotated rx -0.54 ry -0.25 rz -43.22 deg, size 10 x 20 x 5 mm, geometry from box.sld
        - object Box at (557156, 103.35, 13.17) mm, rotated rx -0.53 ry 0.26 rz 8.2 deg, size 10 x 20 x 5 mm, geometry from box.sld
        - object Box at (556484, 103.35, 13.17) mm, rotated rx -0.59 ry -0.05 rz -23.16 deg, size 10 x 20 x 5 mm, geometry from box.sld
        - object Box at (555823, 103.35, 13.17) mm, rotated rx -0.39 ry 0.45 rz 30.79 deg, size 10 x 20 x 5 mm, geometry from box.sld
        - object Box at (555157, 103.35, 13.17) mm, rotated rx -0.53 ry 0.27 rz 9.07 deg, size 10 x 20 x 5 mm, geometry from box.sld
        - object Box at (554486, 103.35, 13.17) mm, rotated rx -0.59 ry -0.02 rz -20.11 deg, size 10 x 20 x 5 mm, geometry from box.sld
        - object Box at (553818, 103.35, 13.17) mm, rotated rx -0.59 ry -0.01 rz -18.86 deg, size 10 x 20 x 5 mm, geometry from box.sld
        - object Box at (553143, 103.35, 13.17) mm, rotated rx -0.41 ry 0.43 rz 28.32 deg, size 10 x 20 x 5 mm, geometry from box.sld
        - object Box at (552476, 103.35, 13.17) mm, rotated rx -0.59 ry 0.02 rz -16.39 deg, size 10 x 20 x 5 mm, geometry from box.sld
        - object Box at (551799, 103.35, 13.17) mm, rotated rx -0.59 ry -0.09 rz -26.42 deg, size 10 x 20 x 5 mm, geometry from box.sld
        - object Box at (551127, 103.35, 13.17) mm, rotated rx -0.42 ry 0.42 rz 27.39 deg, size 10 x 20 x 5 mm, geometry from box.sld
        - object Box at (550461, 103.35, 13.17) mm, rotated rx -0.55 ry 0.22 rz 3.26 deg, size 10 x 20 x 5 mm, geometry from box.sld
        - object Box at (549789, 103.35, 13.17) mm, rotated rx -0.57 ry 0.16 rz -2.57 deg, size 10 x 20 x 5 mm, geometry from box.sld
        - object Box at (549118, 103.35, 13.17) mm, rotated rx -0.59 ry 0 rz -18.42 deg, size 10 x 20 x 5 mm, geometry from box.sld
        - object Box at (548442, 103.35, 13.17) mm, rotated rx -0.53 ry 0.27 rz 8.4 deg, size 10 x 20 x 5 mm, geometry from box.sld
        - object Box at (547768, 103.35, 13.17) mm, rotated rx -0.57 ry 0.16 rz -2.27 deg, size 10 x 20 x 5 mm, geometry from box.sld
        - object Box at (547097, 103.35, 13.17) mm, rotated rx -0.59 ry 0.09 rz -9.8 deg, size 10 x 20 x 5 mm, geometry from box.sld
        - object Box at (546420, 103.35, 13.17) mm, rotated rx -0.48 ry 0.35 rz 18.52 deg, size 10 x 20 x 5 mm, geometry from box.sld
        - object Box at (545744, 103.35, 13.17) mm, rotated rx -0.37 ry 0.47 rz 33.7 deg, size 10 x 20 x 5 mm, geometry from box.sld
        - object Box at (545061, 103.35, 13.17) mm, rotated rx -0.46 ry 0.38 rz 21.15 deg, size 10 x 20 x 5 mm, geometry from box.sld
        - object Box at (544387, 103.35, 13.17) mm, rotated rx -0.47 ry 0.36 rz 18.82 deg, size 10 x 20 x 5 mm, geometry from box.sld
        - object Box at (543712, 103.35, 13.17) mm, rotated rx -0.48 ry 0.35 rz 18.29 deg, size 10 x 20 x 5 mm, geometry from box.sld
        - object Box at (543029, 103.35, 13.17) mm, rotated rx -0.5 ry 0.32 rz 14.37 deg, size 10 x 20 x 5 mm, geometry from box.sld
        - object Box at (542348, 103.35, 13.17) mm, rotated rx -0.58 ry -0.13 rz -30.82 deg, size 10 x 20 x 5 mm, geometry from box.sld
        - object Box at (541667, 103.35, 13.17) mm, rotated rx -0.57 ry 0.16 rz -2.06 deg, size 10 x 20 x 5 mm, geometry from box.sld
        - object Box at (540975, 103.35, 13.17) mm, rotated rx -0.56 ry 0.2 rz 1.42 deg, size 10 x 20 x 5 mm, geometry from box.sld
        - object Box at (540296, 103.35, 13.17) mm, rotated rx -0.56 ry 0.2 rz 1.38 deg, size 10 x 20 x 5 mm, geometry from box.sld
        - object Box at (539623, 103.35, 13.17) mm, rotated rx -0.39 ry 0.44 rz 30.17 deg, size 10 x 20 x 5 mm, geometry from box.sld
        - object Box at (538944, 103.35, 13.17) mm, rotated rx -0.58 ry 0.1 rz -8.26 deg, size 10 x 20 x 5 mm, geometry from box.sld
        - object Box at (538267, 103.35, 13.17) mm, rotated rx -0.59 ry -0.01 rz -19.06 deg, size 10 x 20 x 5 mm, geometry from box.sld
        - object Box at (537589, 103.35, 13.17) mm, rotated rx -0.59 ry -0.05 rz -23.05 deg, size 10 x 20 x 5 mm, geometry from box.sld
        - object Box at (536912, 103.35, 13.17) mm, rotated rx -0.58 ry 0.14 rz -4.62 deg, size 10 x 20 x 5 mm, geometry from box.sld
        - object Box at (536231, 103.35, 13.17) mm, rotated rx -0.59 ry 0.08 rz -10.27 deg, size 10 x 20 x 5 mm, geometry from box.sld
        - object Box at (535546, 103.35, 13.17) mm, rotated rx -0.51 ry 0.3 rz 12.04 deg, size 10 x 20 x 5 mm, geometry from box.sld
        - object Box at (534871, 103.35, 13.17) mm, rotated rx -0.59 ry -0.07 rz -25.12 deg, size 10 x 20 x 5 mm, geometry from box.sld
        - object Box at (534189, 103.35, 13.17) mm, rotated rx -0.58 ry 0.12 rz -6.55 deg, size 10 x 20 x 5 mm, geometry from box.sld
        - object Box at (533505, 103.35, 13.17) mm, rotated rx -0.59 ry 0.08 rz -10.76 deg, size 10 x 20 x 5 mm, geometry from box.sld
        - object Box at (532826, 103.35, 13.17) mm, rotated rx -0.5 ry 0.32 rz 14.46 deg, size 10 x 20 x 5 mm, geometry from box.sld
        - object Box at (532144, 103.35, 13.17) mm, rotated rx -0.56 ry 0.21 rz 2.14 deg, size 10 x 20 x 5 mm, geometry from box.sld
        - object Box at (531464, 103.35, 13.17) mm, rotated rx -0.59 ry -0.03 rz -21.02 deg, size 10 x 20 x 5 mm, geometry from box.sld
        - object Box at (530781, 103.35, 13.17) mm, rotated rx -0.59 ry 0.06 rz -11.91 deg, size 10 x 20 x 5 mm, geometry from box.sld
        - object Box at (530096, 103.35, 13.17) mm, rotated rx -0.38 ry 0.46 rz 32.64 deg, size 10 x 20 x 5 mm, geometry from box.sld
        - object Box at (529411, 103.35, 13.17) mm, rotated rx -0.36 ry 0.47 rz 34.89 deg, size 10 x 20 x 5 mm, geometry from box.sld
        - object Box at (528729, 103.35, 13.17) mm, rotated rx -0.58 ry 0.11 rz -7.78 deg, size 10 x 20 x 5 mm, geometry from box.sld
        - object Box at (528046, 103.35, 13.17) mm, rotated rx -0.57 ry 0.17 rz -1.12 deg, size 10 x 20 x 5 mm, geometry from box.sld
        - object Box at (527361, 103.35, 13.17) mm, rotated rx -0.39 ry 0.45 rz 30.98 deg, size 10 x 20 x 5 mm, geometry from box.sld
        - object Box at (526672, 103.35, 13.17) mm, rotated rx -0.46 ry 0.38 rz 21.54 deg, size 10 x 20 x 5 mm, geometry from box.sld
        - object Box at (525986, 103.35, 13.17) mm, rotated rx -0.59 ry 0.02 rz -16.1 deg, size 10 x 20 x 5 mm, geometry from box.sld
        - object Box at (525299, 103.35, 13.17) mm, rotated rx -0.58 ry -0.13 rz -31.12 deg, size 10 x 20 x 5 mm, geometry from box.sld
        - object Box at (524613, 103.35, 13.17) mm, rotated rx -0.59 ry 0.03 rz -15.33 deg, size 10 x 20 x 5 mm, geometry from box.sld
        - object Box at (523928, 103.35, 13.17) mm, rotated rx -0.59 ry 0.09 rz -9.78 deg, size 10 x 20 x 5 mm, geometry from box.sld
        - object Box at (523238, 103.35, 13.17) mm, rotated rx -0.53 ry -0.27 rz -44.88 deg, size 10 x 20 x 5 mm, geometry from box.sld
        - object Box at (522545, 103.35, 13.17) mm, rotated rx -0.59 ry 0.08 rz -10.21 deg, size 10 x 20 x 5 mm, geometry from box.sld
        - object Box at (521859, 103.35, 13.17) mm, rotated rx -0.58 ry -0.11 rz -28.5 deg, size 10 x 20 x 5 mm, geometry from box.sld
        - object Box at (521172, 103.35, 13.17) mm, rotated rx -0.41 ry 0.43 rz 28.72 deg, size 10 x 20 x 5 mm, geometry from box.sld
        - object Box at (520487, 103.35, 13.17) mm, rotated rx -0.47 ry 0.36 rz 18.77 deg, size 10 x 20 x 5 mm, geometry from box.sld
        - object Box at (519788, 103.35, 13.17) mm, rotated rx -0.31 ry 0.51 rz 40.15 deg, size 10 x 20 x 5 mm, geometry from box.sld
        - object Box at (519098, 103.35, 13.17) mm, rotated rx -0.59 ry 0.1 rz -8.75 deg, size 10 x 20 x 5 mm, geometry from box.sld
        - object Box at (518411, 103.35, 13.17) mm, rotated rx -0.48 ry 0.35 rz 18.27 deg, size 10 x 20 x 5 mm, geometry from box.sld
        - object Box at (517721, 103.35, 13.17) mm, rotated rx -0.59 ry -0.09 rz -26.57 deg, size 10 x 20 x 5 mm, geometry from box.sld
        - object Box at (517027, 103.35, 13.17) mm, rotated rx -0.59 ry -0.09 rz -26.46 deg, size 10 x 20 x 5 mm, geometry from box.sld
        - object Box at (516333, 103.35, 13.17) mm, rotated rx -0.37 ry 0.46 rz 33.17 deg, size 10 x 20 x 5 mm, geometry from box.sld
        - object Box at (515640, 103.35, 13.17) mm, rotated rx -0.59 ry 0.06 rz -12.21 deg, size 10 x 20 x 5 mm, geometry from box.sld
        - object Box at (514947, 103.35, 13.17) mm, rotated rx -0.55 ry -0.22 rz -40 deg, size 10 x 20 x 5 mm, geometry from box.sld
        - object Box at (514253, 103.35, 13.17) mm, rotated rx -0.59 ry 0.02 rz -15.81 deg, size 10 x 20 x 5 mm, geometry from box.sld
        - object Box at (513563, 103.35, 13.17) mm, rotated rx -0.59 ry -0.06 rz -23.81 deg, size 10 x 20 x 5 mm, geometry from box.sld
        - object Box at (512875, 103.35, 13.17) mm, rotated rx -0.54 ry -0.24 rz -41.94 deg, size 10 x 20 x 5 mm, geometry from box.sld
        - object Box at (512182, 103.35, 13.17) mm, rotated rx -0.54 ry 0.25 rz 7.03 deg, size 10 x 20 x 5 mm, geometry from box.sld
        - object Box at (511486, 103.35, 13.17) mm, rotated rx -0.58 ry 0.14 rz -4.94 deg, size 10 x 20 x 5 mm, geometry from box.sld
        - object Box at (510791, 103.35, 13.17) mm, rotated rx -0.43 ry 0.41 rz 25.22 deg, size 10 x 20 x 5 mm, geometry from box.sld
        - object Box at (510098, 103.35, 13.17) mm, rotated rx -0.58 ry 0.13 rz -5.7 deg, size 10 x 20 x 5 mm, geometry from box.sld
        - object Box at (509398, 103.35, 13.17) mm, rotated rx -0.59 ry -0.07 rz -25.18 deg, size 10 x 20 x 5 mm, geometry from box.sld
        - object Box at (508703, 103.35, 13.17) mm, rotated rx -0.43 ry 0.4 rz 24.82 deg, size 10 x 20 x 5 mm, geometry from box.sld
        - object Box at (508008, 103.35, 13.17) mm, rotated rx -0.31 ry 0.51 rz 40.19 deg, size 10 x 20 x 5 mm, geometry from box.sld
        - object Box at (507295, 103.35, 13.17) mm, rotated rx -0.58 ry 0.12 rz -6.59 deg, size 10 x 20 x 5 mm, geometry from box.sld
        - object Box at (506604, 103.35, 13.17) mm, rotated rx -0.59 ry -0.08 rz -25.96 deg, size 10 x 20 x 5 mm, geometry from box.sld
        - object Box at (505904, 103.35, 13.17) mm, rotated rx -0.51 ry 0.31 rz 13.31 deg, size 10 x 20 x 5 mm, geometry from box.sld
        - object Box at (505203, 103.35, 13.17) mm, rotated rx -0.59 ry -0.08 rz -26.26 deg, size 10 x 20 x 5 mm, geometry from box.sld
        - object Box at (504480, 103.35, 13.17) mm, rotated rx -0.59 ry 0 rz -18.1 deg, size 10 x 20 x 5 mm, geometry from box.sld
        - object Box at (503778, 103.35, 13.17) mm, rotated rx -0.45 ry 0.39 rz 22.8 deg, size 10 x 20 x 5 mm, geometry from box.sld
        - object Box at (503071, 103.35, 13.17) mm, rotated rx -0.59 ry -0.01 rz -18.96 deg, size 10 x 20 x 5 mm, geometry from box.sld
        - object Box at (502366, 103.35, 13.17) mm, rotated rx -0.59 ry 0.06 rz -11.96 deg, size 10 x 20 x 5 mm, geometry from box.sld
        - object Box at (501664, 103.35, 13.17) mm, rotated rx -0.5 ry 0.31 rz 13.68 deg, size 10 x 20 x 5 mm, geometry from box.sld
        - object Box at (500959, 103.35, 13.17) mm, rotated rx -0.36 ry 0.47 rz 34.25 deg, size 10 x 20 x 5 mm, geometry from box.sld
        - object Box at (500263, 103.35, 13.17) mm, rotated rx -0.52 ry 0.28 rz 9.83 deg, size 10 x 20 x 5 mm, geometry from box.sld
        - object Box at (499608, 103.35, 13.17) mm, rotated rx -0.57 ry -0.18 rz -35.63 deg, size 10 x 20 x 5 mm, geometry from box.sld
        - object Box at (498912, 103.35, 13.17) mm, rotated rx -0.57 ry -0.17 rz -34.9 deg, size 10 x 20 x 5 mm, geometry from box.sld
        - object Box at (498210, 103.35, 13.17) mm, rotated rx -0.59 ry -0.01 rz -19.6 deg, size 10 x 20 x 5 mm, geometry from box.sld
        - object Box at (497504, 103.35, 13.17) mm, rotated rx -0.59 ry 0.04 rz -14.42 deg, size 10 x 20 x 5 mm, geometry from box.sld
        - object Box at (496806, 103.35, 13.17) mm, rotated rx -0.59 ry -0.09 rz -26.58 deg, size 10 x 20 x 5 mm, geometry from box.sld
        - object Box at (496102, 103.35, 13.17) mm, rotated rx -0.55 ry 0.22 rz 3.88 deg, size 10 x 20 x 5 mm, geometry from box.sld
        - object Box at (495401, 103.35, 13.17) mm, rotated rx -0.29 ry 0.52 rz 42.07 deg, size 10 x 20 x 5 mm, geometry from box.sld
        - object Box at (494688, 103.35, 13.17) mm, rotated rx -0.27 ry 0.53 rz 44.31 deg, size 10 x 20 x 5 mm, geometry from box.sld
        - object Box at (493983, 103.35, 13.17) mm, rotated rx -0.56 ry 0.19 rz 0.89 deg, size 10 x 20 x 5 mm, geometry from box.sld
        - object Box at (493281, 103.35, 13.17) mm, rotated rx -0.59 ry 0.06 rz -12.63 deg, size 10 x 20 x 5 mm, geometry from box.sld
        - object Box at (492575, 103.35, 13.17) mm, rotated rx -0.59 ry -0.04 rz -22.21 deg, size 10 x 20 x 5 mm, geometry from box.sld
        - object Box at (491864, 103.35, 13.17) mm, rotated rx -0.57 ry 0.16 rz -2.39 deg, size 10 x 20 x 5 mm, geometry from box.sld
        - object Box at (491159, 103.35, 13.17) mm, rotated rx -0.59 ry -0.07 rz -25.15 deg, size 10 x 20 x 5 mm, geometry from box.sld
        - object Box at (490455, 103.35, 13.17) mm, rotated rx -0.45 ry 0.39 rz 22.48 deg, size 10 x 20 x 5 mm, geometry from box.sld
        - object Box at (489748, 103.35, 13.17) mm, rotated rx -0.36 ry 0.47 rz 34.83 deg, size 10 x 20 x 5 mm, geometry from box.sld
        - object Box at (489045, 103.35, 13.17) mm, rotated rx -0.33 ry 0.49 rz 37.5 deg, size 10 x 20 x 5 mm, geometry from box.sld
        - object Box at (488339, 103.35, 13.17) mm, rotated rx -0.58 ry 0.13 rz -5.2 deg, size 10 x 20 x 5 mm, geometry from box.sld
        - object Box at (487628, 103.35, 13.17) mm, rotated rx -0.31 ry 0.51 rz 40.7 deg, size 10 x 20 x 5 mm, geometry from box.sld
        - object Box at (486922, 103.35, 13.17) mm, rotated rx -0.57 ry -0.16 rz -34.2 deg, size 10 x 20 x 5 mm, geometry from box.sld
        - object Box at (486216, 103.35, 13.17) mm, rotated rx -0.29 ry 0.52 rz 42.61 deg, size 10 x 20 x 5 mm, geometry from box.sld
        - object Box at (485502, 103.35, 13.17) mm, rotated rx -0.58 ry 0.1 rz -8.36 deg, size 10 x 20 x 5 mm, geometry from box.sld
        - object Box at (484790, 103.35, 13.17) mm, rotated rx -0.58 ry -0.12 rz -30.12 deg, size 10 x 20 x 5 mm, geometry from box.sld
        - object Box at (484077, 103.35, 13.17) mm, rotated rx -0.39 ry 0.45 rz 30.51 deg, size 10 x 20 x 5 mm, geometry from box.sld
        - object Box at (483365, 103.35, 13.17) mm, rotated rx -0.58 ry 0.12 rz -6.95 deg, size 10 x 20 x 5 mm, geometry from box.sld
        - object Box at (482651, 103.35, 13.17) mm, rotated rx -0.59 ry 0.05 rz -12.88 deg, size 10 x 20 x 5 mm, geometry from box.sld
        - object Box at (481942, 103.35, 13.17) mm, rotated rx -0.34 ry 0.49 rz 37.27 deg, size 10 x 20 x 5 mm, geometry from box.sld
        - object Box at (481230, 103.35, 13.17) mm, rotated rx -0.59 ry -0.05 rz -23.22 deg, size 10 x 20 x 5 mm, geometry from box.sld
        - object Box at (480516, 103.35, 13.17) mm, rotated rx -0.59 ry -0.08 rz -25.69 deg, size 10 x 20 x 5 mm, geometry from box.sld
        - object Box at (479804, 103.35, 13.17) mm, rotated rx -0.59 ry -0.01 rz -19.07 deg, size 10 x 20 x 5 mm, geometry from box.sld
        - object Box at (479082, 103.35, 13.17) mm, rotated rx -0.47 ry 0.37 rz 19.92 deg, size 10 x 20 x 5 mm, geometry from box.sld
        - object Box at (478374, 103.35, 13.17) mm, rotated rx -0.56 ry -0.21 rz -38.53 deg, size 10 x 20 x 5 mm, geometry from box.sld
        - object Box at (477664, 103.35, 13.17) mm, rotated rx -0.56 ry 0.19 rz 0.96 deg, size 10 x 20 x 5 mm, geometry from box.sld
        - object Box at (476948, 103.35, 13.17) mm, rotated rx -0.42 ry 0.42 rz 26.27 deg, size 10 x 20 x 5 mm, geometry from box.sld
        - object Box at (476238, 103.35, 13.17) mm, rotated rx -0.3 ry 0.51 rz 41.02 deg, size 10 x 20 x 5 mm, geometry from box.sld
        - object Box at (475500, 103.35, 13.17) mm, rotated rx -0.55 ry -0.22 rz -39.51 deg, size 10 x 20 x 5 mm, geometry from box.sld
        - object Box at (474793, 103.35, 13.17) mm, rotated rx -0.35 ry 0.48 rz 35.67 deg, size 10 x 20 x 5 mm, geometry from box.sld
        - object Box at (474076, 103.35, 13.17) mm, rotated rx -0.57 ry -0.15 rz -32.77 deg, size 10 x 20 x 5 mm, geometry from box.sld
        - object Box at (473358, 103.35, 13.17) mm, rotated rx -0.38 ry 0.46 rz 32.55 deg, size 10 x 20 x 5 mm, geometry from box.sld
        - object Box at (472639, 103.35, 13.17) mm, rotated rx -0.59 ry -0.07 rz -25.11 deg, size 10 x 20 x 5 mm, geometry from box.sld
        - object Box at (471919, 103.35, 13.17) mm, rotated rx -0.56 ry -0.19 rz -36.43 deg, size 10 x 20 x 5 mm, geometry from box.sld
        - object Box at (471203, 103.35, 13.17) mm, rotated rx -0.59 ry -0.08 rz -25.54 deg, size 10 x 20 x 5 mm, geometry from box.sld
        - object Box at (470486, 103.35, 13.17) mm, rotated rx -0.55 ry -0.23 rz -40.97 deg, size 10 x 20 x 5 mm, geometry from box.sld
        - object Box at (469768, 103.35, 13.17) mm, rotated rx -0.39 ry 0.44 rz 30.13 deg, size 10 x 20 x 5 mm, geometry from box.sld
        - object Box at (469058, 103.35, 13.17) mm, rotated rx -0.55 ry 0.22 rz 3.22 deg, size 10 x 20 x 5 mm, geometry from box.sld
        - object Box at (468341, 103.35, 13.17) mm, rotated rx -0.59 ry -0.02 rz -19.62 deg, size 10 x 20 x 5 mm, geometry from box.sld
        - object Box at (467571, 103.35, 13.17) mm, rotated rx -0.59 ry 0.07 rz -11.34 deg, size 10 x 20 x 5 mm, geometry from box.sld
        - object Box at (466804, 103.35, 13.17) mm, rotated rx -0.59 ry 0.05 rz -13.65 deg, size 10 x 20 x 5 mm, geometry from box.sld
        - object Box at (466021, 103.35, 13.17) mm, rotated rx -0.51 ry 0.31 rz 12.8 deg, size 10 x 20 x 5 mm, geometry from box.sld
        - object Box at (465242, 103.35, 13.17) mm, rotated rx -0.59 ry 0 rz -18.56 deg, size 10 x 20 x 5 mm, geometry from box.sld
        - object Box at (464468, 103.35, 13.17) mm, rotated rx -0.57 ry 0.16 rz -2.56 deg, size 10 x 20 x 5 mm, geometry from box.sld
        - object Box at (463708, 103.35, 13.17) mm, rotated rx -0.56 ry 0.19 rz 0.82 deg, size 10 x 20 x 5 mm, geometry from box.sld
        - object Box at (462911, 103.35, 13.17) mm, rotated rx -0.51 ry 0.31 rz 13.05 deg, size 10 x 20 x 5 mm, geometry from box.sld
        - object Box at (462136, 103.35, 13.17) mm, rotated rx -0.46 ry 0.38 rz 21.33 deg, size 10 x 20 x 5 mm, geometry from box.sld
        - object Box at (461354, 103.35, 13.17) mm, rotated rx -0.5 ry 0.32 rz 14.26 deg, size 10 x 20 x 5 mm, geometry from box.sld
        - object Box at (460585, 103.35, 13.17) mm, rotated rx -0.53 ry 0.26 rz 8.2 deg, size 10 x 20 x 5 mm, geometry from box.sld
        - object Box at (459795, 103.35, 13.17) mm, rotated rx -0.54 ry 0.25 rz 7.2 deg, size 10 x 20 x 5 mm, geometry from box.sld
        - object Box at (459015, 103.35, 13.17) mm, rotated rx -0.37 ry 0.46 rz 33.25 deg, size 10 x 20 x 5 mm, geometry from box.sld
        - object Box at (458219, 103.35, 13.17) mm, rotated rx -0.47 ry 0.37 rz 20.03 deg, size 10 x 20 x 5 mm, geometry from box.sld
        - object Box at (457444, 103.35, 13.17) mm, rotated rx -0.56 ry 0.18 rz -0.24 deg, size 10 x 20 x 5 mm, geometry from box.sld
        - object Box at (456652, 103.35, 13.17) mm, rotated rx -0.33 ry 0.49 rz 37.97 deg, size 10 x 20 x 5 mm, geometry from box.sld
        - object Box at (455877, 103.35, 13.17) mm, rotated rx -0.55 ry 0.22 rz 3.59 deg, size 10 x 20 x 5 mm, geometry from box.sld
        - object Box at (455092, 103.35, 13.17) mm, rotated rx -0.58 ry 0.12 rz -6.01 deg, size 10 x 20 x 5 mm, geometry from box.sld
        - object Box at (454337, 103.35, 13.17) mm, rotated rx -0.54 ry 0.24 rz 6.17 deg, size 10 x 20 x 5 mm, geometry from box.sld
        - object Box at (453547, 103.35, 13.17) mm, rotated rx -0.56 ry -0.2 rz -38.29 deg, size 10 x 20 x 5 mm, geometry from box.sld
        - object Box at (452765, 103.35, 13.17) mm, rotated rx -0.53 ry 0.27 rz 8.84 deg, size 10 x 20 x 5 mm, geometry from box.sld
        - object Box at (451977, 103.35, 13.17) mm, rotated rx -0.34 ry 0.48 rz 36.63 deg, size 10 x 20 x 5 mm, geometry from box.sld
        - object Box at (451197, 103.35, 13.17) mm, rotated rx -0.59 ry 0.01 rz -16.83 deg, size 10 x 20 x 5 mm, geometry from box.sld
        - object Box at (450421, 103.35, 13.17) mm, rotated rx -0.55 ry 0.23 rz 4.68 deg, size 10 x 20 x 5 mm, geometry from box.sld
        - object Box at (449644, 103.35, 13.17) mm, rotated rx -0.58 ry -0.14 rz -31.98 deg, size 10 x 20 x 5 mm, geometry from box.sld
        - object Box at (448866, 103.35, 13.17) mm, rotated rx -0.4 ry 0.43 rz 28.82 deg, size 10 x 20 x 5 mm, geometry from box.sld
        - object Box at (448089, 103.35, 13.17) mm, rotated rx -0.57 ry 0.16 rz -2.47 deg, size 10 x 20 x 5 mm, geometry from box.sld
        - object Box at (447300, 103.35, 13.17) mm, rotated rx -0.59 ry 0 rz -18.37 deg, size 10 x 20 x 5 mm, geometry from box.sld
        - object Box at (446517, 103.35, 13.17) mm, rotated rx -0.38 ry 0.46 rz 32.13 deg, size 10 x 20 x 5 mm, geometry from box.sld
        - object Box at (445740, 103.35, 13.17) mm, rotated rx -0.57 ry 0.17 rz -1.03 deg, size 10 x 20 x 5 mm, geometry from box.sld
        - object Box at (444967, 103.35, 13.17) mm, rotated rx -0.59 ry 0.03 rz -15.58 deg, size 10 x 20 x 5 mm, geometry from box.sld
        - object Box at (444175, 103.35, 13.17) mm, rotated rx -0.49 ry 0.34 rz 16.87 deg, size 10 x 20 x 5 mm, geometry from box.sld
        - object Box at (443402, 103.35, 13.17) mm, rotated rx -0.42 ry 0.42 rz 27.01 deg, size 10 x 20 x 5 mm, geometry from box.sld
        - object Box at (442616, 103.35, 13.17) mm, rotated rx -0.31 ry 0.5 rz 39.89 deg, size 10 x 20 x 5 mm, geometry from box.sld
        - object Box at (441839, 103.35, 13.17) mm, rotated rx -0.5 ry 0.33 rz 15.25 deg, size 10 x 20 x 5 mm, geometry from box.sld
        - object Box at (441033, 103.35, 13.17) mm, rotated rx -0.58 ry 0.14 rz -4.95 deg, size 10 x 20 x 5 mm, geometry from box.sld
        - object Box at (440247, 103.35, 13.17) mm, rotated rx -0.46 ry 0.37 rz 20.91 deg, size 10 x 20 x 5 mm, geometry from box.sld
        - object Box at (439434, 103.35, 13.17) mm, rotated rx -0.57 ry -0.17 rz -35.29 deg, size 10 x 20 x 5 mm, geometry from box.sld
        - object Box at (438642, 103.35, 13.17) mm, rotated rx -0.59 ry 0.04 rz -14.42 deg, size 10 x 20 x 5 mm, geometry from box.sld
        - object Box at (437838, 103.35, 13.17) mm, rotated rx -0.57 ry -0.17 rz -34.74 deg, size 10 x 20 x 5 mm, geometry from box.sld
